(* IEC 61131-3 sources: SortJet_MasterSPS_Aufbau.fbsproj/09_Station/Shuttle/[101,102] Shuttle, 9 files *)

(* ---- Dickenverstellung_FB_V01_00_00.fb.st ---- *)
(* METADATA
{
	"v3Meta": {
		"objectGuid": "d815e3f2-dcd5-4a25-9c13-c3ee247e2cce"
	}
}
*)
FUNCTION_BLOCK Dickenverstellung_FB_V01_00_00
VAR_INPUT

  // BOOLEAN
  bpAktivieren                                   : BOOL; // Hinweis: Baustein aktivieren
  bpReset                                        : BOOL;
  bpStartePositionierung                         : BOOL;
  bpReferenz                                     : BOOL;
  bpFreigabe                                     : BOOL;
  bpOptionMotorischAktivieren                    : BOOL;
  bpOptionPneumatikAktivieren                    : BOOL;
  bpOption3WegeLogikDrehen                       : BOOL;
  bpOptionRollenleisteSchuetzSchaltungAktivieren : BOOL;
  bpOptionGegenhalterSchuetzSchaltungAktivieren  : BOOL;

  // ENUM
  epSollStellung : PneumatikZylinderStatus_EN;

  // STRUCT
  stStationsNummern  : Station_ST;

  // POINTER
  ppAntriebsInformationen : REFERENCE TO AntriebsInformationen;
  ppParameterBaustein     : REFERENCE TO Parameter_Dickenverstellung;  // Zeiger auf Parameterfeld

END_VAR
VAR_OUTPUT

  // BOOLEAN
  bpFehler                  : BOOL;
  bpDone                    : BOOL;
  bpResourceAktiv           : BOOL;
  bpInReferenz              : BOOL; // Status: Baustein/Antrieb ist referenziert

  // WORD
  wpFehlerNr : Fehlerkonstanten_EN;

  // ENUM
  eStatusStellung : PneumatikZylinderStatus_EN;

END_VAR
VAR

  // BOOLEAN
  blErsterZyklus   : BOOL := TRUE;

  // REAL
  rlZielPosition   : REAL;

  // TIMER
  tonlEndschalterFreifahren              : TON; // EINSCHALTVERZOEGERUNG:
  tonlWarteSchrittEndschalterFreifahren  : TON; // EINSCHALTVERZOEGERUNG:
  tonlMaxWarteAufResetErfolgreich        : TON; // EINSCHALTVERZOEGERUNG:
  tofHardwareEndschalterFrei             : TOF; // AUSSCHALTVERZOEGERUNG:
  toflAutoAbschaltung                    : TOF; // AUSSCHALTVERZOEGERUNG:

  // STEPS
  steplPositionieren    : Steps_TE;
  steplReferenz         : Steps_TE;
  steplReset            : Steps_TE;

  // Antrieb
  Antrieb : REFERENCE TO Rexroth_ctrlX_Drive_Eckelmann_MC_V01_02_02;

END_VAR
VAR_INPUT

  // HARDWARE EINGAENGE
  in_bEndschalterMax : BOOL; // Oeffner (TRUE = frei), gemappt; zum Umrichter ueber Signal-Steuerwort Bit 9, wirkt nur bei Endschalterquelle SPS

END_VAR
//-------------------------------------------------------------------------------------------------
// INITIALISIERUNG
//-------------------------------------------------------------------------------------------------
IF ( blErsterZyklus ) THEN

  IF ( __ISVALIDREF(ppAntriebsInformationen) ) THEN

    blErsterZyklus := FALSE;

    Antrieb REF= pgAntriebe[ppAntriebsInformationen.wAchsID];

    (* Hinweis:
       - Initialisierung Antriebsinformationen
    *)
    Antrieb.ppAntriebsInformationen REF= ppAntriebsInformationen;

    (* Hinweis:
       - Für die Zielpunktkontrolle muss im ersten Zyklus die Zielposition initialisiert werden
    *)
    Antrieb.rpZielPosition := Antrieb.rpIstPosition;

    (* Hinweis:
       - Antriebswerte vorinitialisieren
    *)
    Antrieb.rpGeschwindigkeit := ppAntriebsInformationen.rpMaxGeschwindigkeit;
    Antrieb.rpBeschleunigung  := ppAntriebsInformationen.rpMaxBeschleunigung;
    Antrieb.rpVerzoegerung    := ppAntriebsInformationen.rpMaxVerzoegerung;
    Antrieb.rpRuckzeit        := ppAntriebsInformationen.rpMaxRuckzeit;

  ELSE
    RETURN;
  END_IF

END_IF

// Endschalter zyklisch an den Antrieb geben, auch bei deaktivierter Bewegung
Antrieb.bpEndschalterMaxExtern := in_bEndschalterMax;

//-------------------------------------------------------------------------------------------------
// BAUSTEIN: AUSFUEHRUNG
//-------------------------------------------------------------------------------------------------
(* Hinweis:
   - Aktionen
*)
IF ( bpReset AND bpAktivieren ) THEN

  Reset();

ELSE

  IF ( bpAktivieren ) THEN
    Positionieren();
    Referenz();
    Ausgaenge();

    (* Hinweis:
       - Abschaltung
    *)
    toflAutoAbschaltung( IN :=     bpStartePositionierung
                         OR bpReferenz,
                         PT:= tgZeitAutoabschaltungEnergiesparModus );

    Antrieb.bpFreigabe := toflAutoAbschaltung.Q
                          AND bpAktivieren
                          AND bpFreigabe;

    Antrieb.rpRuckzeit := ppAntriebsInformationen.rpMaxRuckzeit;

    Antrieb.stStationsNummern := stStationsNummern;

  ELSE
    bpDone   := TRUE;
    bpFehler := FALSE;
    bpInReferenz := TRUE;

    eStatusStellung := epSollStellung;

    wpFehlerNr := cMELDUNG_NULL;

  END_IF // => bpAktiv

END_IF// => bpReset
END_FUNCTION_BLOCK

(* ---- Dickenverstellung_Schuetz_FB_V01_00_00.fb.st ---- *)
(* METADATA
{
	"v3Meta": {
		"objectGuid": "2c7452d1-eabd-4c4a-95fd-5aca04df1ee1"
	}
}
*)
FUNCTION_BLOCK Dickenverstellung_Schuetz_FB_V01_00_00
VAR_INPUT

  // BOOL
  bpAktivieren               : BOOL;
  bpVerstellungOeffnen       : BOOL;
  bpVerstellungSchliessen    : BOOL;
  bpReset                    : BOOL;

END_VAR
VAR_OUTPUT

  // BOOL
  bpFehler        : BOOL;
  bpDone          : BOOL;
  bpResourceAktiv : BOOL;

  // WORD
  wpFehlerNr      : Fehlerkonstanten_EN;

END_VAR

VAR

  // BOOL
  blErsterZyklus        : BOOL := TRUE;

  // TIMER
  tonlMaxWarteZeit                        : TON;
  tonlAntriebOK                           : TON;
  tonlMaximaleWartezeitAufReset           : TON;
  tonlFehlermeldungUnterdrueckenAntriebOK : TON;

  // STEPS
  steplVerstellungOeffnen      : Steps_TE;
  steplVerstellungSchliessen   : Steps_TE;
  steplReset                   : Steps_TE;

END_VAR

VAR
  // HARDWARE EINGÄNGE
  in_bVerstellungGeoeffnet         AT %I* : BOOL;
  in_bVerstellungGeschlossen       AT %I* : BOOL;
  in_bMotorstarter_OK              AT %I* : BOOL; // Sicherung des Kippantriebs ÖFFNER KONTAKT !!
  in_bBremseOK                     AT %I* : BOOL; // Sicherung des Kippantriebs ÖFFNER KONTAKT !!
  in_bSicherungMotorOK             AT %I* : BOOL;

  // HARDWARE AUSGÄNGE
  out_bVerstellungSchliessen       AT %Q* : BOOL;
  out_bVerstellungOeffnen          AT %Q* : BOOL;
  out_bBremseOeffnen               AT %Q* : BOOL;
  out_bMotorstarterReset           AT %Q* : BOOL;

END_VAR

//-------------------------------------------------------------------------------------------------
// BAUSTEIN: INITIALISIERUNG
//-------------------------------------------------------------------------------------------------
IF ( blErsterZyklus ) THEN
  blErsterZyklus := FALSE;

  (* Hinweis:
     - Timer initialisieren
  *)
  tonlAntriebOK(IN:=TRUE);
  tonlMaxWarteZeit(IN:=FALSE);
  tonlFehlermeldungUnterdrueckenAntriebOK( IN := FALSE );

END_IF

//-------------------------------------------------------------------------------------------------
// BAUSTEIN: AKTIONEN
//-------------------------------------------------------------------------------------------------
(* Hinweis:
   - Aktionen
*)
IF ( bpReset ) THEN

  bpReset                 := FALSE;
  bpVerstellungOeffnen    := FALSE;
  bpVerstellungSchliessen := FALSE;

  bpFehler        := FALSE;
  bpDone          := FALSE;
  bpResourceAktiv := FALSE;

  wpFehlerNr := cMELDUNG_NULL;

  out_bVerstellungSchliessen  := FALSE;
  out_bVerstellungOeffnen := FALSE;

ELSE

  IF ( bpAktivieren ) THEN

    VerstellungSchliessen();
    VerstellungOeffnen();

    out_bBremseOeffnen := out_bVerstellungOeffnen OR out_bVerstellungSchliessen;

    Meldungen();
    Timer();

  ELSE

    bpDone   := TRUE;
    bpFehler := FALSE;

  END_IF // => bpAktiv

END_IF// => bpReset
END_FUNCTION_BLOCK

(* ---- Greiferzange_FB_V01_00_00.fb.st ---- *)
(* METADATA
{
	"v3Meta": {
		"objectGuid": "50b45b59-5893-4c9c-b524-1732205d1fb3"
	}
}
*)
FUNCTION_BLOCK Greiferzange_FB_V01_00_00
VAR_INPUT

  // BOOLEAN
  bpReset                     : BOOL;
  bpAktivieren                : BOOL;
  bpFreigabe                  : BOOL; // FREIGABE Pneumatik: ohne Freigabe Ventile aus, Bewegung pausiert (Startbefehl bleibt erhalten)
  bpStartZylinderBewegung     : BOOL; // BETRIEBTYP: Greiferzange in die Soll-Stellung bewegen
  bpZylinderAbfragenVorhanden : BOOL := FALSE; // Hinweis: Endlagenabfragen der Zylinder vorhanden

  // TIME
  tpBewegungszeit             : TIME := T#700MS; // Bewegungszeit je Stellung ohne Abfragen bzw. beim Schliessen auf Glas

  // ENUM
  epSollZylinderStellung      : PneumatikZylinderStatus_EN; // eZylinderGeschlossen, eZylinderStellung16mm, eZylinderStellung23mm, eZylinderStellung29mm

END_VAR
VAR_OUTPUT

  // BOOLEAN
  bpFehler                    : BOOL;
  bpDone                      : BOOL;

  // WORD
  wpFehlerNr                  : Fehlerkonstanten_EN;

  // ENUM
  epStatusZylinderStellung    : PneumatikZylinderStatus_EN;

END_VAR
VAR

  // STEPS
  steplZylinderStellung       : Steps_TE;

  // TIMER
  tonlUeberwachungStellung      : TON; // EINSCHALTVERZOEGERUNG: Ueberwachung der Soll-Stellung mit Abfragen
  tonlWartezeitZylinderStellung : TON; // EINSCHALTVERZOEGERUNG: Bewegungszeit ohne Abfragen

END_VAR
VAR

  // HARDWARE EINGAENGE
  in_bStatusZylinder_Alle_Eingefahren AT %I* : BOOL; // STATUS: Zylinderabfrage [Eingefahren] Zange geschlossen
  in_bStatusZylinder_1_Ausgefahren    AT %I* : BOOL; // STATUS: Zylinderabfrage [Ausgefahren] Oeffnung 16 mm
  in_bStatusZylinder_2_Ausgefahren    AT %I* : BOOL; // STATUS: Zylinderabfrage [Ausgefahren] Oeffnung 23 mm
  in_bStatusZylinder_3_Ausgefahren    AT %I* : BOOL; // STATUS: Zylinderabfrage [Ausgefahren] Oeffnung 29 mm

  // HARDWARE AUSGAENGE
  out_bZylinder_1_Einfahren           AT %Q* : BOOL; // Impuls Zylinder 1 einfahren
  out_bZylinder_2_Einfahren           AT %Q* : BOOL; // Impuls Zylinder 2 einfahren
  out_bZylinder_3_Einfahren           AT %Q* : BOOL; // Impuls Zylinder 3 einfahren
  out_bZylinder_1_Ausfahren           AT %Q* : BOOL; // Impuls Zylinder 1 ausfahren [16 mm]
  out_bZylinder_2_Ausfahren           AT %Q* : BOOL; // Impuls Zylinder 2 ausfahren [23 mm]
  out_bZylinder_3_Ausfahren           AT %Q* : BOOL; // Impuls Zylinder 3 ausfahren [29 mm]

END_VAR
VAR CONSTANT

  // TIME
  cZEIT_UEBERWACHUNG_STELLUNG : TIME := T#5S;

END_VAR
(* Anmerkung:
   - Greiferzange mit drei Zylindern: geschlossen, Oeffnung 16 mm, 23 mm oder 29 mm
   - Vor dem Oeffnen werden alle Zylinder eingefahren, danach faehrt der Zylinder der Soll-Oeffnung aus
*)
//-------------------------------------------------------------------------------------------------
// BAUSTEIN: RESET / DEAKTIVIERT
//-------------------------------------------------------------------------------------------------
(* Hinweis:
   - Reset oder deaktiviert: Ausgaenge aus, Kette und Timer zuruecksetzen, Done und Fehler loeschen
   - Der Baustein setzt bpReset selbst zurueck, der Aufrufer wartet nicht auf Done
   - Ein deaktivierter Baustein meldet kein Done; der Aufrufer verknuepft das Warten auf Done
     mit der Aktivierung aus der MK (z.B. Greiferzange.bpDone OR NOT stStationsAufbau.bGreifer[wWand])
*)
IF ( bpReset OR NOT bpAktivieren ) THEN

  out_bZylinder_1_Einfahren := FALSE;
  out_bZylinder_2_Einfahren := FALSE;
  out_bZylinder_3_Einfahren := FALSE;
  out_bZylinder_1_Ausfahren := FALSE;
  out_bZylinder_2_Ausfahren := FALSE;
  out_bZylinder_3_Ausfahren := FALSE;

  bpStartZylinderBewegung := FALSE;

  steplZylinderStellung := STEP_0_E;

  tonlUeberwachungStellung( IN := FALSE );
  tonlWartezeitZylinderStellung( IN := FALSE );

  bpDone     := FALSE;
  bpFehler   := FALSE;
  wpFehlerNr := cMELDUNG_NULL;

  bpReset := FALSE;

  RETURN;

END_IF

//-------------------------------------------------------------------------------------------------
// BAUSTEIN: AKTIONEN
//-------------------------------------------------------------------------------------------------
(* Hinweis Freigabe Pneumatik:
   - Ohne Freigabe: Ventile aus, Kette und Ueberwachungszeiten zuruecksetzen (kein Timeout-Fehler)
   - Der Startbefehl bleibt erhalten: kommt die Freigabe zurueck, wird die Bewegung neu gestartet
*)
IF NOT bpFreigabe THEN
  out_bZylinder_1_Einfahren := FALSE;
  out_bZylinder_2_Einfahren := FALSE;
  out_bZylinder_3_Einfahren := FALSE;
  out_bZylinder_1_Ausfahren := FALSE;
  out_bZylinder_2_Ausfahren := FALSE;
  out_bZylinder_3_Ausfahren := FALSE;
  steplZylinderStellung := STEP_0_E;
  tonlUeberwachungStellung( IN := FALSE );
  tonlWartezeitZylinderStellung( IN := FALSE );
  bpDone := FALSE;
ELSE
  ZylinderBewegung();
END_IF

//-------------------------------------------------------------------------------------------------
// STATUS DER ZYLINDER
//-------------------------------------------------------------------------------------------------
(* Hinweis:
   - Status aus der Sensorik, wenn Abfragen vorhanden sind
   - Ohne Abfragen bleibt der Status, den die Schrittkette nach der Bewegungszeit setzt
*)
IF ( bpZylinderAbfragenVorhanden ) THEN

  IF ( in_bStatusZylinder_3_Ausgefahren ) THEN
    epStatusZylinderStellung := eZylinderStellung29mm;

  ELSIF ( in_bStatusZylinder_2_Ausgefahren ) THEN
    epStatusZylinderStellung := eZylinderStellung23mm;

  ELSIF ( in_bStatusZylinder_1_Ausgefahren ) THEN
    epStatusZylinderStellung := eZylinderStellung16mm;

  ELSIF ( in_bStatusZylinder_Alle_Eingefahren ) THEN
    epStatusZylinderStellung := eZylinderGeschlossen;

  ELSE
    epStatusZylinderStellung := eZylinderUndefiniert;

  END_IF

END_IF
END_FUNCTION_BLOCK

(* ---- Shuttle_FB_V01_00_00.fb.st ---- *)
(* METADATA
{
	"v3Meta": {
		"objectGuid": "a8175c8a-0e5e-42c5-a90c-c5e1a843dc34"
	}
}
*)
FUNCTION_BLOCK Shuttle_FB_V01_00_00
VAR_IN_OUT

  // STRUKT
  BasisStationsParameter : StationBasisParameter_ST;

END_VAR
VAR_INPUT

  // BOOLEAN
  bpShuttleAnhalten                      : BOOL; // HINWEIS: Nehmen der Verfahrfreigabe wenn bei der Folge- bzw. Nachfolgestation der Einlauf- / Auslauf- Sensor belegt wurde
  bpStarteFaecherwagensuche              : BOOL; // Der Fächerwagen kann mittels Sensor gesucht werden um die Fachpositionen zu bestimmen

  // WORD
  rpMinPosSwEsEingrenzung                : REAL;
  rpMaxPosSwEsEingrenzung                : REAL;

END_VAR
VAR_OUTPUT

  // BOOLEAN
  bpFaecherwagenGefunden                 : BOOL;

  // REAL
  rpAktuelleFaecherwagenPosition         : REAL;

  // DWORD
  dwpHandfunktionenReturn                : DWORD; // Aktive Handfunktionen, gleiche Bitbelegung wie dwlHandfunktionen

END_VAR
VAR

  // BOOL
  blErsterZyklus                         : BOOL := TRUE;// Initialisierungsphase
  blGeblaeseAktiv                        : BOOL;
  blBetriebsartHand                      : BOOL;
  blBetriebsartReset                     : BOOL;
  blBetriebartCheck                      : BOOL;
  blBetriebsartAutomatik                 : BOOL;
  blBetriebsartReferenz                  : BOOL;
  ablZielPositionErreicht                : ARRAY[cWAND_1..cANZAHL_WAENDE] OF BOOL; // Je Wand: Zielposition aus dem Auftrag der Wand stimmt mit der aktuellen Position ueberein [Toleranz rgMKZielPositionToleranz]
  blVorAbAuftragAktiv                    : ARRAY [cWAND_1..cANZAHL_WAENDE] OF BOOL; // STATUS: Merker ob die Komponenten Ansteuerung aktiv ist [Angesteuert mit dem Starten der Querfahrt](Autark gesteuert)
  blUpdateTimer                          : BOOL;
  blNachSystemcheckMerker                : BOOL; // Merkt sich, wenn der Systemcheck erfolgreich durchgeführt wurde, damit die Gebläse nicht nach dem Systemcheck ausgehen
  ablVortransportAktiv                   : ARRAY [cWAND_1..cANZAHL_WAENDE] OF BOOL; // STATUS: Merker ob der Vortransport (Autark gesteuert) aktiv ist -> Wichtig für den Austransport zum sicherstellen das erst dann Transportiert werden kann
  blDatenlichtschrankeUnterbrochenMelden : BOOL;
  blFehlerAusAutomatikBetrieb            : BOOL;
  blShuttleErreichbar                    : BOOL;
  blMerkerAuftragAktiv                   : BOOL;
  blMerkerEinOderAustransportAktiv       : BOOL;

  // WORD
  wlBetriebsart              : WORD;
  wlWatchIONachrichtenNummer : WORD;
  wlIndex                    : WORD;

  // DWORD
  dwlHandfunktionen                : DWORD;  // Handfunktionen: 0..31 Bit
  dwlHandfunktionenZuletztGesendet : DWORD;  // Rueckmeldung der Handfunktionen zum MMI

  // REAL
  rlLetztePosition  : REAL;

  // TIMER
  tonlMaxWarteAufResetErfolgreich       : TON;
  tonlUpdateTimer                       : TON; // Verfahrlogik
  tonWaitTimerAnsteuerungResourcen      : ARRAY[cWAND_1..cANZAHL_WAENDE] OF TON;
  tonWaitTimerAnsteuerungResourcenDone  : ARRAY[cWAND_1..cANZAHL_WAENDE] OF TON;

  toflGeblaeseHandfahren                : ARRAY[cWAND_1..cANZAHL_WAENDE] OF TOF;
  atoflSensorEinlauf                    : ARRAY[cWAND_1..cANZAHL_WAENDE] OF TOF;
  atoflSensorAuslauf                    : ARRAY[cWAND_1..cANZAHL_WAENDE] OF TOF;
  atoflSensorAUslaufStopp               : ARRAY[cWAND_1..cANZAHL_WAENDE] OF TOF;
  atoflSensorEinlaufStopp               : ARRAY[cWAND_1..cANZAHL_WAENDE] OF TOF;

  // TRIGGER
  rtlAutomatikActiv                     : R_TRIG;
  rtlGlastransportVerfahrfreigabe       : ARRAY [cWAND_1..cANZAHL_WAENDE] OF R_TRIG;
  rtlDatenlichtschrankeUnterbrochen     : R_TRIG;
  rtlFehlerMeldungGenerierenHandbetrieb : R_TRIG;
  rtlFehlerAusgeloestImAutomatikbetrieb : R_TRIG;
  artlVerfahrabbruchSensorik            : ARRAY [cWAND_1..cANZAHL_WAENDE] OF R_TRIG;
  artlWandverstellungPositionieren      : ARRAY [cWAND_1..cANZAHL_WAENDE] OF R_TRIG;
  rtlRackPositionGefunden               : R_TRIG;
  ftlBausteinDeaktivierung              : F_TRIG;

  // STEPS
  steplCheck                       : STEPS_TE;
  steplResetAntrieb                : STEPS_TE;
  steplReferenz                    : Steps_TE;
  steplVorabpositionierung         : STEPS_TE;
  steplFaecherwagensuche           : STEPS_TE;

  // BAUSTEINE
  Querfahrt                       : Querfahrt_Shuttle_FB_V01_00_00;
  Zentralschmierung               : Zentralschmierung_DLS_4xxi_FB_V01_00_00;
  Glastransport                   : ARRAY[cWAND_1..cANZAHL_WAENDE] OF Shuttle_Glastransport_FB_V01_00_00;
  Geblaese                        : ARRAY[cWAND_1..cANZAHL_WAENDE] OF Geblaese_Schuetz_FB_V01_00_00;
  Wandverstellung                 : ARRAY[cWAND_1..cANZAHL_WAENDE] OF Dickenverstellung_FB_V01_00_00;
  Kippen                          : Shuttle_Kippen_V01_00_00;

  Eintransport                    : ARRAY[cWAND_1..cANZAHL_WAENDE] OF Shuttle_Eintransport_FB_V01_00_00;
  Austransport                    : ARRAY[cWAND_1..cANZAHL_WAENDE] OF Shuttle_Austransport_FB_V01_00_00;
  Durchtransport                  : ARRAY[cWAND_1..cANZAHL_WAENDE] OF Shuttle_Durchtransport_FB_V01_00_00;
  AnsteuerungRessourcen           : ARRAY[cWAND_1..cANZAHL_WAENDE] OF Shuttle_Ansteuerung_Ressourcen_FB_V01_00_00;
  Greifer                         : ARRAY[cWAND_1..cANZAHL_WAENDE] OF Shuttle_Greifer_FB_V01_00_00; // Ausbaustufe stStationsAufbau.bGreifer

END_VAR
VAR
  // Alle Sensoren
  blAlleEinlaufStoppSensoren : BOOL; // wirksame Einlauf-Stopp-Sensoren (ohne MK: Einlaufsensor)
  blAlleAuslaufStoppSensoren : BOOL;
  ablSensorEinlaufStopp      : ARRAY[cWAND_1..cANZAHL_WAENDE] OF BOOL; // wirksamer Einlauf-Stopp-Sensor (ohne MK: Einlaufsensor)
  ablSensorAuslaufStopp      : ARRAY[cWAND_1..cANZAHL_WAENDE] OF BOOL; // wirksamer Auslauf-Stopp-Sensor (ohne MK: Auslaufsensor)
  blAlleVerfahrfreigaben     : BOOL;
  blAlleGreiferSicher        : BOOL; // Alle Greifer in sicherer Position mit eingefahrenen Glasrueckhaltern (oder nicht vorhanden)
  blGreiferVor               : BOOL; // Handbetrieb Greifer: Taster MMI oder Visu (Aktion Handfunktionen)
  blGreiferZurueck           : BOOL;
  blGreiferReferenz          : BOOL;
  blGreiferAusfahren         : BOOL;
  blGreiferEinfahren         : BOOL;
  ablQuittScheibe            : ARRAY[cWAND_1..cANZAHL_WAENDE] OF BOOL; // Scheibenquittierung Glastransport bzw. Greifer
  blDone                     : BOOL;
  blFehlerAktiv              : BOOL;

  // HARDWARE EINGAENGE
  in_bSensorEinlauf                                   : ARRAY[cWAND_1..cANZAHL_WAENDE] OF BOOL; // Shuttle Sensoren von links nach rechts Sensor 1
  in_bSensorAuslauf                                   : ARRAY[cWAND_1..cANZAHL_WAENDE] OF BOOL; // Shuttle Sensoren von links nach rechts Sensor 4
  in_bSensorEinlaufVorab                              : ARRAY[cWAND_1..cANZAHL_WAENDE] OF BOOL; // Shuttle Sensoren von links nach rechts Sensor 2
  in_bSensorAuslaufVorab                              : ARRAY[cWAND_1..cANZAHL_WAENDE] OF BOOL; // Shuttle Sensoren von links nach rechts Sensor 3
  in_bSensorEinlaufStopp                              : ARRAY[cWAND_1..cANZAHL_WAENDE] OF BOOL; // Shuttle Sensoren von links nach rechts Sensor 0 (nur mit MK bSensorEinlaufStopp)
  in_bSensorAuslaufStopp                              : ARRAY[cWAND_1..cANZAHL_WAENDE] OF BOOL; // Shuttle Sensoren von links nach rechts Sensor 5 (nur mit MK bSensorAuslaufStopp)
  in_bDatenlichtschrankeShuttlebahnOK          AT %I* : BOOL; // Bauteil an der Shuttlebahn => Sender / Empfaenger
  in_bDatenlichtschrankeShuttleOK              AT %I* : BOOL; // Bauteil auf dem Shuttle => Sender / Empfaenger
  in_bNetzteil_24V_OK                          AT %I* : BOOL;
  in_bKlimageraet_OK                                  : BOOL;
  in_bSicherungen24V_OK                               : BOOL;
  in_bDruckluft_OK                             AT %I* : BOOL;
  in_bSicherungKompressor_OK                   AT %I* : BOOL;
  in_bLSQuerfahrtBremseOK                      AT %I* : BOOL;

  in_bSicherungen230V_OK                       AT %I* : BOOL;
  in_iAnalogwertChannel1                              : INT; // Hinweis: Eingaenge des Analogmoduls u.a fuer die automatische Fachaufnahme
  in_iAnalogwertChannel2                              : INT; // Hinweis: Eingaenge des Analogmoduls u.a fuer die automatische Fachaufnahme
  in_bWandverstellungsAntriebsSicherungOK      AT %I* : BOOL;
  in_bWandverstellungsBremsSicherungOK         AT %I* : BOOL;
  in_bFaecherwagenSuchSensor                          : BOOL; // Shuttle Sensor zum Suchen der Fächerwagen um die Fachpositionen zu bestimmen

  aHand : ARRAY[0..31] OF BOOL;
  i     : INT;

END_VAR
VAR CONSTANT

  // TIME
  ZEIT_SENSOR_ENTPRELLEN         : TIME := T#50ms;

END_VAR
(* Anmerkung:
   - Shuttle Koordinationsbaustein regelt das komplette Shuttle
*)
//-------------------------------------------------------------------------------------------------
// BAUSTEIN: INITIALISIERUNG
//-------------------------------------------------------------------------------------------------

IF ( blErsterZyklus ) THEN
  blErsterZyklus:=FALSE;

  (* Wichtig:
     - Initialisierung
  *)
  A_Baustein_Initialisierung();

END_IF

FOR wlIndex := cWAND_1 TO cANZAHL_WAENDE DO
  in_bSensorEinlauf[wlIndex] := Glastransport[wlIndex].Antrieb.udipEingaengeUmrichter.cXG31_1_I_1;
  in_bSensorAuslauf[wlIndex] := Glastransport[wlIndex].Antrieb.udipEingaengeUmrichter.cXG31_2_I_2;

  ablSensorEinlaufStopp[wlIndex] := SEL( BasisStationsParameter.stMKs.stStationsAufbau.bSensorEinlaufStopp, in_bSensorEinlauf[wlIndex], in_bSensorEinlaufStopp[wlIndex] );
  ablSensorAuslaufStopp[wlIndex] := SEL( BasisStationsParameter.stMKs.stStationsAufbau.bSensorAuslaufStopp, in_bSensorAuslauf[wlIndex], in_bSensorAuslaufStopp[wlIndex] );
END_FOR

blAlleEinlaufStoppSensoren := FALSE;
blAlleAuslaufStoppSensoren := FALSE;
blAlleVerfahrfreigaben     := TRUE;
blAlleGreiferSicher        := TRUE;

FOR wlIndex := cWAND_1 TO cANZAHL_WAENDE DO
  blAlleGreiferSicher        := blAlleGreiferSicher
                                AND (    ( Greifer[wlIndex].bpSicherePosition AND Greifer[wlIndex].bpGlasRueckhalterEingefahren )
                                      OR NOT BasisStationsParameter.stMKs.stStationsAufbau.bGreifer[wlIndex] );
  blAlleEinlaufStoppSensoren := blAlleEinlaufStoppSensoren OR ablSensorEinlaufStopp[wlIndex];
  blAlleAuslaufStoppSensoren := blAlleAuslaufStoppSensoren OR ablSensorAuslaufStopp[wlIndex];
  blAlleVerfahrfreigaben     := blAlleVerfahrfreigaben AND Glastransport[wlIndex].bpVerfahrFreigabe;
END_FOR

//-------------------------------------------------------------------------------------------------
// DEAKTIVIERUNG
//-------------------------------------------------------------------------------------------------

(* Hinweis:
   - Werte wieder passend abloeschen, wenn der Baustein wieder aktiviert wird
*)
ftlBausteinDeaktivierung( CLK := BasisStationsParameter.stMKs.bDeaktivieren );

IF ( ftlBausteinDeaktivierung.Q ) THEN

  SendShuttlePosition();

  FOR wlIndex := cWAND_1 TO cANZAHL_WAENDE DO
    BasisStationsParameter.bEintransportAbgeschlossen[wlIndex] := FALSE;
    BasisStationsParameter.bAustransportAbgeschlossen[wlIndex] := FALSE;
  END_FOR

  BasisStationsParameter.bIstReferenziert       := FALSE;
  BasisStationsParameter.bCheckAbgeschlossen    := FALSE;
  BasisStationsParameter.bReferenzAbgeschlossen := FALSE;

END_IF

(* Hinweis:
   - Deaktivierung des Bausteins
     => Der Baustein wird zum Ende der RETURN-Anweisung verlassen
*)
IF ( BasisStationsParameter.stMKs.bDeaktivieren ) THEN

  IF ( apgShuttleVerfahrparameter[BasisStationsParameter.stMKs.stStationsNummern.NummerSPS].eParkposition = PARKPOSITION_MAX ) THEN
    BasisStationsParameter.rAktuellePositionQuerfahrt := apgShuttleVerfahrparameter[BasisStationsParameter.stMKs.stStationsNummern.NummerSPS].rParkpositionMaximum;
  ELSE
    BasisStationsParameter.rAktuellePositionQuerfahrt := apgShuttleVerfahrparameter[BasisStationsParameter.stMKs.stStationsNummern.NummerSPS].rParkpositionMinimum;
  END_IF

  FOR wlIndex := cWAND_1 TO cANZAHL_WAENDE DO
    BasisStationsParameter.bEintransportAbgeschlossen[wlIndex] := TRUE;
    BasisStationsParameter.bAustransportAbgeschlossen[wlIndex] := TRUE;

    IF ( BasisStationsParameter.bCheck ) THEN

      IF BasisStationsParameter.stMKs.stStationsAufbau.bGlastransport[wlIndex] THEN
        rSps2MmiMessungScheibenlaenge   := 0;
        wSps2MmiMessungStationNummer    := BasisStationsParameter.stMKs.stStationsNummern.NummerIntern;
        wSps2MmiMessungSlotNummer       := wlIndex;
        iSps2MmiMessungScheibenanzahl   := 0;

        MsgToMmi( auftragsnr_w := SB0_SPS_SETSHEETSONSTATION );
      END_IF
    END_IF

  END_FOR

  BasisStationsParameter.bIstReferenziert       := TRUE;
  BasisStationsParameter.bCheckAbgeschlossen    := TRUE;
  BasisStationsParameter.bReferenzAbgeschlossen := TRUE;
  BasisStationsParameter.bReset                 := FALSE;

  BasisStationsParameter.bFehler       := FALSE;
  BasisStationsParameter.wFehlerNummer := cMELDUNG_NULL;

  HandfunktionenStatus();
  RETURN;

END_IF

//-------------------------------------------------------------------------------------------------
// AKTIONEN
//-------------------------------------------------------------------------------------------------
Betriebsart();

SystemCheck();

(* Hinweis:
   - Automatik-Aktionen
*)
FOR wlIndex := cWAND_1 TO cANZAHL_WAENDE DO
  Eintransport[wlIndex]( BasisStationsParameter := BasisStationsParameter,
                         wWand := wlIndex,
                         bpGeblaeseAktiv := Geblaese[wlIndex].bpDone,
                         bpAutomatikAktiv := BasisStationsParameter.bAutomatik,
                         bpVorAbAuftragAktiv := blVorAbAuftragAktiv[wlIndex],
                         bpZielPositionErreicht := ablZielPositionErreicht[wlIndex],
                         Glastransport := Glastransport[wlIndex],
                         Kippen := Kippen,
                         Wandverstellung := Wandverstellung[wlIndex],
                         Geblaese := Geblaese[wlIndex],
                         bpGreiferAktiv := BasisStationsParameter.stMKs.stStationsAufbau.bGreifer[wlIndex],
                         Greifer := Greifer[wlIndex]
                       );
  Austransport[wlIndex]( BasisStationsParameter := BasisStationsParameter,
                         wWand := wlIndex,
                         bpGeblaeseAktiv := Geblaese[wlIndex].bpDone,
                         bpAutomatikAktiv := BasisStationsParameter.bAutomatik,
                         bpVorAbAuftragAktiv := blVorAbAuftragAktiv[wlIndex],
                         bpZielPositionErreicht := ablZielPositionErreicht[wlIndex],
                         Glastransport := Glastransport[wlIndex],
                         Kippen := Kippen,
                         Wandverstellung := Wandverstellung[wlIndex],
                         Geblaese := Geblaese[wlIndex],
                         bpGreiferAktiv := BasisStationsParameter.stMKs.stStationsAufbau.bGreifer[wlIndex],
                         Greifer := Greifer[wlIndex]
                       );

  Durchtransport[wlIndex]( BasisStationsParameter := BasisStationsParameter,
                           wWand := wlIndex,
                           bpGeblaeseAktiv := Geblaese[wlIndex].bpDone,
                           bpAutomatikAktiv := BasisStationsParameter.bAutomatik,
                           bpVorAbAuftragAktiv := blVorAbAuftragAktiv[wlIndex],
                           bpZielPositionErreicht := ablZielPositionErreicht[wlIndex],
                           Glastransport := Glastransport[wlIndex],
                           Kippen := Kippen,
                           Wandverstellung := Wandverstellung[wlIndex],
                           Geblaese := Geblaese[wlIndex]
                         );
  AnsteuerungRessourcen[wlIndex]( BasisStationsParameter := BasisStationsParameter,
                                  wWand := wlIndex,
                                  bpGeblaeseAktiv := Geblaese[wlIndex].bpDone,
                                  bpAutomatikAktiv := BasisStationsParameter.bAutomatik,
                                  bpVorAbAuftragAktiv := blVorAbAuftragAktiv[wlIndex],
                                  bpZielPositionErreicht := ablZielPositionErreicht[wlIndex],
                                  Glastransport := Glastransport[wlIndex],
                                  Kippen := Kippen,
                                  Wandverstellung := Wandverstellung[wlIndex],
                                  Geblaese := Geblaese[wlIndex],
                                  bpGreiferAktiv := BasisStationsParameter.stMKs.stStationsAufbau.bGreifer[wlIndex],
                                  Greifer := Greifer[wlIndex]
                                );
END_FOR

Vorabpositionierung();

SensorenFreifahren();
FaecherwagenSuche();

(* Hinweis:
   - Basis-Aktionen
*)
Reset();
Referenz();
Meldungen();
Handfunktionen();

A_Geblaese();
A_Aufrufe();
A_Schnittstelle();
A_Ausgaenge();
END_FUNCTION_BLOCK

(* ---- Shuttle_Glastransport_FB_V01_00_00.fb.st ---- *)
(* METADATA
{
	"v3Meta": {
		"objectGuid": "bced77b5-e61c-4af0-a672-a0da8c7118bb"
	}
}
*)
FUNCTION_BLOCK Shuttle_Glastransport_FB_V01_00_00
VAR_INPUT

  bpDurchtransport                 : BOOL; // BETRIEBSMODUS[AUTOMATIK]: Eintransport-Schrittkette starten
  bpEintransport                   : BOOL; // BETRIEBSMODUS[AUTOMATIK]: Eintransport-Schrittkette starten
  bpRueckwaertsEintransportieren   : BOOL; // BETRIEBSMODUS[AUTOMATIK]: Eintransport Richtung -Rueckwaerts ueber den Auslaufsensor
  bpAustransport                   : BOOL; // BETRIEBSMODUS[AUTOMATIK]: Autransport-Schrittkette starten
  bpRueckwaertsAustransportieren   : BOOL; // BETRIEBSMODUS[AUTOMATIK]: Austransport Richtung -Rueckwaerts ueber den Einlaufsensor
  bpRueckwaertsSystemcheck         : BOOL;
  bpVortransport                   : BOOL; // BETRIEBSMODUS[AUTOMATIK]: Vortransport-Schrittkette starten
  bpVortransportRueck              : BOOL; // BETRIEBSMODUS[AUTOMATIK]: Vortransport-Schrittkette starten
  bpStarteSensorFreiFahren         : BOOL := FALSE; // BETRIEBSMODUS[AUTOMATIK]:
  bpHandfahrenPlus                 : BOOL; // BETRIEBSMODUS HANDBETRIEB: Im Handbetrieb den Riemen in positive Glasflussrichtung bewegen
  bpHandfahrenMinus                : BOOL; // BETRIEBSMODUS HANDBETRIEB: Im Handbetrieb den Riemen in negative Glasflussrichtung bewegen
  bpFahreReferenz                  : BOOL; // BETRIEBSMODUS: Antrieb referenzieren
  bpStarteVorabPositionierung      : BOOL; // BETRIEBSMODUS Positionieren der Scheibe fuer den Austransport
  bpStarteVorabPositionierungRueckwaertig : BOOL; // BETRIEBSMODUS Positionieren der Scheibe fuer den Austransport rueckwaerts (ueber den Einlaufsensor)
  bpCheck                          : BOOL;
  bpReset                          : BOOL;
  bpCheckMitVorgaenger             : BOOL; // Status: SystemCheck mit der Vorgaenger- Station
  bpCheckMitNachfolger             : BOOL; // Status: SystemCheck mit der Nachfolger- Station
  bpAutomatikAktiv                 : BOOL;
  bpFreigabe                       : BOOL; // Status: Der Riemen ist Freigegeben und kann Prozesse abarbeiten
  bpMessrichtungNegativ            : BOOL := FALSE; // HINWEIS: TRUE = Messrichtung negativ, FALSE = Messrichtung positiv
  bpAktivieren                     : BOOL := TRUE; // WICHTIG: Aktivieren des Bausteins
  bpScheibentrennung               : BOOL := FALSE;
  bpTransferstationTransfershuttle : BOOL := FALSE;
  bpSensorEinlauf                  : BOOL; // Sensoren von links nach rechts Sensor 1
  bpSensorEinlaufVorab             : BOOL; // Sensoren von links nach rechts Sensor 2
  bpSensorAuslaufVorab             : BOOL; // Sensoren von links nach rechts Sensor 3
  bpSensorAuslauf                  : BOOL; // Sensoren von links nach rechts Sensor 4
  bpSensorEinlaufStopp             : BOOL; // Sensoren von links nach rechts Sensor 0 (Verfahrfreigabe, Notbremse und Scheibe hat Shuttle verlassen im Rueckwaertstransport)
  bpSensorAuslaufStopp             : BOOL; // Sensoren von links nach rechts Sensor 5
  bpScheibeNachSystemcheckAufAuslaufsensor : BOOL;
  bpTeilnehmerErreichbar           : BOOL;
  bpMessungSystemCheckAktiv        : BOOL;
  bpSlaveAntriebVorhanden          : BOOL;

  // OPTIONEN
  bpOptionMasterSlaveTransport     : BOOL;

  // GREIFER
  bpStarteSlaveKopplungGreifer      : BOOL; // BETRIEBSMODUS GREIFER: Glastransport als Slave auf die Greiferachse koppeln
  bpStarteKorrekturfahrt            : BOOL; // BETRIEBSMODUS GREIFER: Sensor der Greiferseite frei fahren (uebergrosse Scheibe / nach dem Austransport)
  bpKorrekturfahrtRueckwaerts       : BOOL; // BETRIEBSMODUS GREIFER: TRUE = Auslaufsensor frei fahren, FALSE = Einlaufsensor frei fahren
  bpStarteGlasPositionierungGreifer : BOOL; // BETRIEBSMODUS GREIFER: Scheibe fuer den Austransport mit dem Greifer positionieren
  bpGlasPositionierungEinlaufseite  : BOOL; // BETRIEBSMODUS GREIFER: TRUE = ueber den Einlaufsensor positionieren, FALSE = ueber den Auslaufsensor
  wpAchsIDGreifer                   : WORD; // Achs-ID der Greiferachse (Master der Kopplung)
  rpWegGlasUebergabeposition        : REAL; // Weg der Scheibe ueber den Sensor der Greiferseite

  // WORD
  wpWandNr                    : WORD;

  // ENUM
  eStationsTyp                 : StationsTyp_EN; // Typ der Station [ Shuttle \ Station \ Faecherwagen \ etc. ]
  wpGlastyp                   : GlasTyp_EN; // AUFTRAGSDATEN : Unterscheidung fuer den Eintransports -> Grosse Scheiben

  // STRUCT
  InGlasTransportNachfolger   : Interface_GlasTransport; // STRUKTUR: Informationen ueber den Aus- Ein- Transport WAND 2
  InGlasTransportVorgaenger   : Interface_GlasTransport; // STRUKTUR: Informationen ueber den Aus- Ein- Transport WAND 2
  pAuftrag                    : Auftragsdaten_ST;        // AUFTRAG: Aktuelle daten zum Auftrag [Laenge, Hoehe, Modelle]
  stStationsNummern           : Station_ST;
  stMasterSlaveConfig         : MasterSlaveConfig_ST;

  // POINTER
  ppParameterBaustein           : REFERENCE TO Parameter_ShuttleGlastransport;
  ppAntriebsInformationen       : REFERENCE TO AntriebsInformationen;
  ppAntriebsInformationenSlave  : REFERENCE TO AntriebsInformationen;

END_VAR
VAR_OUTPUT

  // BOOLEAN
  bpDone                                      : BOOL;
  bpFehler                                    : BOOL;
  bprtScheibe                                 : BOOL;
  bpStationBelegt                             : BOOL;
  bpVerfahrFreigabe                           : BOOL;
  bpVortransportAktiv                         : BOOL; // STATUS: Merker ob der Vortransport (Autark gesteuert) aktiv ist -> Wichtig für den Austransport zum sicherstellen das erst dann Transportiert werden kann
  bpPositionierungAbgeschlossen               : BOOL; // HINWEIS:
  bpOutBereitZumAustransport                  : BOOL;
  bpOutBereitZumEintransport                  : BOOL;
  bpSlaveAktiv                                : BOOL; // STATUS: dem Baustein melden das der Slavebetrieb aktiv ist
  bpFreigabeQuerfahrt                         : BOOL; // HINWEIS: Freigabe setzen das die Querfahrt verfahren kann
  bpAuftragAktiv                              : BOOL;
  bpGreiferSlaveAktiv                         : BOOL; // STATUS: Glastransport ist auf die Greiferachse gekoppelt
  bpKorrekturfahrtAbgeschlossen               : BOOL; // STATUS: Korrekturfahrt fuer den Greifer abgeschlossen
  bpGlasPositionierungGreiferAbgeschlossen    : BOOL; // STATUS: Scheibe fuer den Greifer positioniert

  // WORD
  wpFehlerNr             : Fehlerkonstanten_EN;

  // DWORD
  dwpWartezeit              : DWORD :=0 ;// STATISTIK: Beschreibt die Zeit zwischen Anlegeauftrag und betaetigen des Tasters zum Eintransport

  // REAL
  rpOutGeschwindigkeit        : REAL;
  rlGlasgewicht               : REAL;

END_VAR
VAR

  // BOOLEAN
  blErsterZyklus                              : BOOL := TRUE;
  blSensorFreifahren                          : BOOL;
  blScheibenMerker                            : BOOL; // Merken da eien Scheibe den Auslaufsensor / Einlaufsensor beim Eintransport weiter
  blReduzierteGeschwindigkeit                 : BOOL;
  blAntriebsKopplungAktiv                     : BOOL;
  blStarteSlaveKopplung                       : BOOL;

  // INT
  ilScheibenZaehler  : INT;

  // REAL
  rlScheibenMessungErgebnis         : REAL; // SystemCheck
  rlAntriebIstPositionBeiStart      : REAL;
  rlMaxStreckeErsteScheibe          : REAL; // Max. Weg bis zur ersten Scheibe: Laenge der abgebenden Station, ohne bekannte Laenge die eigene Stationslaenge
  rlStreckeBisZurVerzoegerung       : REAL;
  rlPositionScheibenAnfangErkannt   : REAL;
  rlGeschwindigkeitEintransport     : REAL;
  rlGefahreneStreckeEintransport    : REAL; // Weg-Merker fuer die Strecke die beim Eintransport zurueck gelegt werden muss laut Auftrag

  // STEPS
  steplDurchtransport           : Steps_TE;
  steplEintransport             : Steps_TE;
  steplEintransportRueckwaertig : Steps_TE;
  steplAustransport             : Steps_TE;
  steplAustransportRueckwaertig : Steps_TE;
  steplSlave                    : Steps_TE;
  steplCheck                    : Steps_TE;
  steplReset                    : Steps_TE;
  steplReferenz                 : Steps_TE;
  steplVorabpositionieren       : STEPS_TE; // Hinweis: Positionierung ueber den Auslaufsensor
  steplVorabpositionierenRueckwaertig : STEPS_TE; // Hinweis: Positionierung ueber den Einlaufsensor
  steplSensorFreiFahren         : Steps_TE;
  steplVortransport             : Steps_TE;
  steplVortransportRueckwertig  : Steps_TE;
  steplSlaveGreifer             : Steps_TE;
  steplKorrekturfahrt           : Steps_TE;
  steplGlasPositionierungGreifer : Steps_TE;

  steplCheckMerker : Steps_TE;

  // TIMER
  toflAutoAbschaltung                : TOF; // AUSSCHALTVERZOEGERUNG:
  toflEinlaufsensor                  : TOF; // AUSSCHALTVERZOEGERUNG: Entprellen der Sensoren
  toflAuslaufsensor                  : TOF; // AUSSCHALTVERZOEGERUNG: Entprellen der Sensoren
  toflAuslaufsensorSTOP              : TOF; // AUSSCHALTVERZOEGERUNG: Entprellen der Sensoren
  toflEinlaufsensorSTOP              : TOF; // AUSSCHALTVERZOEGERUNG: Entprellen der Sensoren
  toflEinlaufsensorFrei              : TOF; // AUSSCHALTVERZOEGERUNG: Haelt die positive Flanke des Auslaufsensor eine gewissen Zeit aufrecht ( Freifahren des Sensors )
  toflAuslaufsensorFrei              : TOF; // AUSSCHALTVERZOEGERUNG: Haelt die positive Flanke des Auslaufsensor eine gewissen Zeit aufrecht ( Freifahren des Sensors )
  tonlMaxWarteAufResetErfolgreich    : TON; // EINSCHALTVERZOEGERUNG:
  tonlWarteSchritt                   : TON; // EINSCHALTVERZOEGERUNG:
  tonlAntriebNichtFreigegeben        : TON; // EINSCHALTVERZOEGERUNG:
  tonlUberwachungSlaveAktiv          : TON; // EINSCHALTVERZOEGERUNG:
  tonlSlaveKopplungDeaktiviert       : TON;
  tonlSlaveAntriebNichtFreigegeben   : TON; // Ueberwachung: Master/Slave nicht betriebsbereit
  tonlUeberwachungSlaveGreifer       : TON; // Ueberwachung: Kopplung auf die Greiferachse
  tonlUeberwachungGreiferBetrieb      : TON; // Ueberwachung: Antrieb bereit fuer Korrekturfahrt / Positionierung fuer den Greifer

  // TIME
  tlWarteZeiteAufnahme               : TIME; // STATISTIK: Zeit Ermittlung von evtl. Wartezeiten

  // STRING
  stlLogString    : STRING;

  // Antrieb
  Scheibenmessung  : Scheibenmessung_FB_V01_00_00;

  // Antrieb
  Antrieb       : REFERENCE TO Rexroth_ctrlX_Drive_Eckelmann_MC_V01_02_02;
  Antrieb_Slave : REFERENCE TO Rexroth_ctrlX_Drive_Eckelmann_MC_V01_02_02;

END_VAR
VAR CONSTANT

  // TIME
  cZEIT_UEBERWACHUNG_ANTRIEBSFREIGABE : TIME := T#5S;
  cUEBERWACHUNG_SLAVE_AKTIV           : TIME :=T#1S;

END_VAR

//-------------------------------------------------------------------------------------------------
// INITIALISIERUNG
//-------------------------------------------------------------------------------------------------
IF ( blErsterZyklus ) THEN

  IF ( __ISVALIDREF(ppAntriebsInformationen) ) THEN

    blErsterZyklus            := FALSE;

    Antrieb REF= pgAntriebe[ppAntriebsInformationen.wAchsID];
    IF ( __ISVALIDREF(ppAntriebsInformationenSlave) ) THEN
      Antrieb_Slave REF= pgAntriebe[ppAntriebsInformationenSlave.wAchsID];
    END_IF

    (* Hinweis:
       - Initialisierung Antriebsinformationen
    *)
    Antrieb.ppAntriebsInformationen REF= ppAntriebsInformationen;
    Antrieb.stStationsNummern := stStationsNummern;
    IF ( __ISVALIDREF(Antrieb_Slave) AND __ISVALIDREF(ppAntriebsInformationenSlave) ) THEN
      Antrieb_Slave.ppAntriebsInformationen REF= ppAntriebsInformationenSlave;
      Antrieb_Slave.stStationsNummern := stStationsNummern;
    END_IF

    (* Hinweis:
       - Antriebswerte vorinitialisieren
    *)
    Antrieb.rpGeschwindigkeit := ppAntriebsInformationen.rpMaxGeschwindigkeit;
    Antrieb.rpBeschleunigung  := ppAntriebsInformationen.rpMaxBeschleunigung;
    Antrieb.rpVerzoegerung    := ppAntriebsInformationen.rpMaxVerzoegerung;
    Antrieb.rpRuckzeit        := ppAntriebsInformationen.rpMaxRuckzeit;

    (* Hinweis:
       - Antriebswerte vorinitialisieren
    *)
    IF ( __ISVALIDREF(Antrieb_Slave) AND __ISVALIDREF(ppAntriebsInformationenSlave) ) THEN
      Antrieb_Slave.rpGeschwindigkeit := REAL#0;
      Antrieb_Slave.rpBeschleunigung  := ppAntriebsInformationenSlave.rpMaxBeschleunigung;
      Antrieb_Slave.rpVerzoegerung    := ppAntriebsInformationenSlave.rpMaxVerzoegerung;
      Antrieb_Slave.rpRuckzeit        := ppAntriebsInformationenSlave.rpMaxRuckzeit;
    END_IF

    // Pointer
    //   - Initialisierung zur vermeidung von null Pointerexceptions
    //     => Scheibenmessung
    Scheibenmessung.ppAntriebsInformationen REF= ppAntriebsInformationen;
    Scheibenmessung.ppAntrieb               REF= Antrieb;
    Scheibenmessung.pbpVorstopSensor        REF= bgFALSE;
    Scheibenmessung.pbpEinlaufSensor        REF= bgFALSE;

  ELSE
    RETURN;
  END_IF

END_IF

//-------------------------------------------------------------------------------------------------
// DEAKTIVIEREN
//-------------------------------------------------------------------------------------------------
IF ( NOT bpAktivieren ) THEN

  bpVerfahrFreigabe := TRUE;
  bpDone := TRUE;

  (* Hinweis:
     - Ausnahmesituationen
  *)
  bpFehler   := FALSE;
  wpFehlerNr := cMELDUNG_NULL;

  RETURN;

END_IF

//-------------------------------------------------------------------------------------------------
// TIMER, EINSTELLUNGEN, ETC.
//-------------------------------------------------------------------------------------------------
(* Hinweis:
   - Sensorenflackern
*)
toflEinlaufsensor(IN := bpSensorEinlauf, PT := t#50ms);
toflAuslaufsensor(IN := bpSensorAuslauf, PT := t#50ms);
toflAuslaufsensorSTOP(IN := bpSensorAuslaufStopp, PT := t#50ms);
toflEinlaufsensorSTOP(IN := bpSensorEinlaufStopp, PT := t#50ms);

// TIMER:
//   - Sensorenflackern
//     => Haelt die positive Flanke des Auslaufsensor eine gewissen Zeit aufrecht ( Freifahren des Sensors )
toflAuslaufsensorFrei(IN := bpSensorAuslauf, PT := t#100ms);
toflEinlaufsensorFrei(IN := bpSensorEinlauf, PT := t#100ms);

//-------------------------------------------------------------------------------------------------
// AKTIONEN
//-------------------------------------------------------------------------------------------------

(* Hinweis:
   - SystemCheck - Aktion
*)
SystemCheck();

(* Hinweis:
   - SystemCheck - Aktion
*)
Eintransport();
Eintransport_Rueckwertig();

Durchtransport();

Austransport();
Austransport_Rueckwertig();

GlasVorabPositionierung();
GlasVorabPositionierung_Rueckwaertig();

CASE eStationsTyp OF

  eInputShuttle:
    Vortransport_Inputshuttle();
    Vortransport_Rueckwertig();

  eOutputShuttle:
    Vortransport();
    Vortransport_Rueckwertig();

END_CASE

SensorenFreifahren();

(* Hinweis:
   - Zusammenspiel mit dem Shuttle-Greifer (nur mit stStationsAufbau.bGreifer angefordert)
*)
GlasPositionierungGreifer();
Korrekturfahrt();
SlaveBetriebGreifer();

IF ( bpSlaveAntriebVorhanden ) THEN
  Slave_Antrieb();
ELSE
  blAntriebsKopplungAktiv := TRUE;
END_IF
(* Hinweis:
   - Basis- Aktionen
*)
Reset();
Referenz();
Meldungen();
Handfunktionen();
Ausgaenge();

//-------------------------------------------------------------------------------------------------
// FREIGABEN UND BAUSTEINAUFRUFE
//-------------------------------------------------------------------------------------------------
(* Hinweis:
   - Freigaben des ANtriebs
*)
toflAutoAbschaltung( IN := (  bpAutomatikAktiv
                             AND ( bpEintransport
                                   OR bpRueckwaertsEintransportieren
                                   OR bpDurchtransport
                                   OR bpVortransport
                                   OR bpVortransportRueck
                                   OR bpAustransport
                                   OR bpRueckwaertsAustransportieren
                                   OR bpStarteSensorFreiFahren
                                   OR bpStarteVorabPositionierung
                                   OR bpStarteVorabPositionierungRueckwaertig
                                   OR bpStarteSlaveKopplungGreifer
                                   OR bpStarteKorrekturfahrt
                                   OR bpStarteGlasPositionierungGreifer ) )
                     OR bpCheck
                     OR bpHandfahrenMinus
                     OR bpHandfahrenPlus
                     OR bpFahreReferenz
                     OR bpStarteSlaveKopplungGreifer
                     OR blStarteSlaveKopplung,
                     PT:= tgZeitAutoabschaltungEnergiesparModus );

// Aufruf Antrieb
Antrieb.bpFreigabe        := toflAutoAbschaltung.Q AND bpFreigabe;
Antrieb.stStationsNummern := stStationsNummern;
Antrieb.rpRuckzeit        := ppAntriebsInformationen.rpMaxRuckzeit;

Antrieb_Slave.bpFreigabe        := toflAutoAbschaltung.Q AND bpFreigabe;
Antrieb_Slave.stStationsNummern := stStationsNummern;
Antrieb_Slave.rpRuckzeit        := ppAntriebsInformationenSlave.rpMaxRuckzeit;

// Aufruf Scheibenmessung
Scheibenmessung( stStationsNummern                   := stStationsNummern,
                 ppAntrieb                           := Antrieb,
                 pbpVorstopSensor                    := bpSensorAuslaufVorab,
                 pbpEinlaufSensor                    := bpSensorEinlauf,
                 bpDrehrichtungsumkehrMessung        := bpMessrichtungNegativ,
                 rpMessstrecke                       := ppParameterBaustein.rMessstrecke,
                 ppAntriebsInformationen             := ppAntriebsInformationen,
                 bpAuswahlSensorVorabScheibenmessung := bgFALSE,
                 epGlastyp                           := wpGlastyp,
                 rpFaktorBremswegverlaengern         := 1.6 ) ;
END_FUNCTION_BLOCK

(* ---- Shuttle_Greifer_FB_V01_00_00.fb.st ---- *)
(* METADATA
{
	"v3Meta": {
		"objectGuid": "bb2ac76d-e136-43b9-91b5-1f4b010b201a"
	}
}
*)
FUNCTION_BLOCK Shuttle_Greifer_FB_V01_00_00
VAR_INPUT

  // BOOLEAN
  bpAktivieren                            : BOOL := FALSE; // WICHTIG: Aktivieren des Bausteins (stStationsAufbau.bGreifer)
  bpFreigabe                              : BOOL; // STATUS: Der Greifer ist freigegeben und kann Prozesse abarbeiten
  bpFreigabePneumatik                     : BOOL; // FREIGABE Pneumatik: Greifer-Hub, Greiferzangen, Glasrueckhalter
  bpAutomatikAktiv                        : BOOL;
  bpTeilnehmerErreichbar                  : BOOL;
  bpReset                                 : BOOL;
  bpFahreReferenz                         : BOOL; // BETRIEBSMODUS: Greiferachse referenzieren
  bpCheck                                 : BOOL; // BETRIEBSMODUS: Systemcheck
  bpStartGrundstellungsfahrt              : BOOL; // BETRIEBSMODUS: Grundstellungsfahrt
  bpPositionieren                         : BOOL; // BETRIEBSMODUS: Greifer hinter die Glaskante positionieren (Laenge aus rpGlaslaenge)
  bpStarteVorabPositionierungEintransport : BOOL; // BETRIEBSMODUS: Greifer vor einem Eintransport an die Wandseite stellen
  bpStarteEintransport                    : BOOL; // BETRIEBSMODUS: Scheibe aus dem Faecherwagen auf das Shuttle ziehen
  bpStarteAustransport                    : BOOL; // BETRIEBSMODUS: Scheibe vom Shuttle in den Faecherwagen schieben
  bpSlaveKopplungAktiv                    : BOOL; // STATUS: Glastransport ist auf die Greiferachse gekoppelt
  bpKorrekturfahrtBeendet                 : BOOL; // STATUS: Korrekturfahrt des Glastransports bei uebergrosser Scheibe abgeschlossen
  bpSensorEinlauf                         : BOOL; // STATUS: Einlaufsensor
  bpSensorAuslauf                         : BOOL; // STATUS: Auslaufsensor

  // HANDBETRIEB
  bpHandfahrenPlus                        : BOOL; // Greiferachse in positive Richtung
  bpHandfahrenMinus                       : BOOL; // Greiferachse in negative Richtung
  bpHandGreiferAusfahren                  : BOOL;
  bpHandGreiferEinfahren                  : BOOL;
  bpHandZangeSchliessen                   : BOOL;
  bpHandZangeOeffnen16mm                  : BOOL;
  bpHandZangeOeffnen23mm                  : BOOL;
  bpHandZangeOeffnen29mm                  : BOOL;
  bpHandGlasRueckhalterAusfahren          : BOOL;

  // ENUM
  epGreiferTyp                            : Greifertyp_EN; // AUFTRAGSDATEN: Greiferseite, eGreiferDefault = Seite aus der MK

  // REAL
  rpGlaslaenge                            : REAL; // Scheibenlaenge fuer das Positionieren hinter die Glaskante

  // STRUCT
  pAuftrag                                : Auftragsdaten_ST; // AUFTRAG: Aktuelle Daten zum Auftrag [Laenge, Hoehe, Dicke, Zangenstellung]
  stStationsNummern                       : Station_ST;

  // POINTER
  ppParameterGreifer                      : REFERENCE TO Parameter_Greifer;
  ppAntriebsInformationen                 : REFERENCE TO AntriebsInformationen;

END_VAR
VAR_OUTPUT

  // BOOLEAN
  bpDone                                         : BOOL; // Reset bzw. Referenz abgeschlossen
  bpFehler                                       : BOOL;
  bprtScheibe                                    : BOOL; // Scheibe quittieren
  bpIstInReferenz                                : BOOL;
  bpSicherePosition                              : BOOL; // WICHTIG: Greifer ragt nicht ueber das Shuttle -> Querfahrt erlaubt
  bpGlasRueckhalterEingefahren                   : BOOL; // WICHTIG: Glasrueckhalter eingefahren -> Querfahrt erlaubt
  bpAnforderungSlaveKopplung                     : BOOL; // Anforderung: Glastransport auf die Greiferachse koppeln
  bpKorrekturfahrtAnfordern                      : BOOL; // Anforderung: Glastransport zieht den Rest einer uebergrossen Scheibe auf das Shuttle
  bpKorrekturfahrtRueckwaerts                    : BOOL; // Richtung der Korrekturfahrt: Sensor der Greiferseite frei fahren
  bpAuftragAktiv                                 : BOOL;
  bpVorpositioniertEintransport                  : BOOL; // Greifer steht ausgefahren an der Wandseite fuer den Eintransport
  bpPositionierungAbgeschlossen                  : BOOL;
  bpVorabPositionierungEintransportAbgeschlossen : BOOL;
  bpEintransportAbgeschlossen                    : BOOL;
  bpAustransportAbgeschlossen                    : BOOL;
  bpGrundstellungsfahrtAbgeschlossen             : BOOL;
  bpSystemCheckAbgeschlossen                     : BOOL;

  // WORD
  wpFehlerNr                                     : Fehlerkonstanten_EN;
  wpFehlerKennung                                : WORD; // Zylinder-Kennung bei Zylinderfehlern (cZYLINDER_*), sonst cZYLINDER_KEINE
  awpFehlerInformationen                        : ARRAY[0..25] OF WORD;

  // REAL
  rpWegGlasUebergabeposition                     : REAL; // Weg der Scheibe ueber den Sensor der Greiferseite vor dem Austransport
  rpIstPosition                                  : REAL;

  // ENUM
  epGreiferTypAktiv                              : Greifertyp_EN; // Greiferseite, mit der gearbeitet wird

END_VAR
VAR

  // BOOLEAN
  blErsterZyklus              : BOOL := TRUE;
  blReduzierteGeschwindigkeit : BOOL;
  blUebergrosseScheibe        : BOOL; // Scheibe zu lang, um sie komplett mit dem Greifer zu ziehen
  blSensorSeite               : BOOL; // Sensor der Greiferseite
  blSensorGegenseite          : BOOL; // Sensor der gegenueberliegenden Seite
  blHandAktiv                 : BOOL;
  blZangeSeiteVorhanden       : BOOL; // Greiferzange der aktiven Greiferseite laut MK vorhanden
  blCheckScheibeZiehen        : BOOL; // Systemcheck: Scheibe im Greifer wird auf das Shuttle gezogen (sonst in den Faecherwagen geschoben)
  blCheckNichtQuittieren      : BOOL; // Systemcheck: Greiferzange war offen, die Scheibe wird nicht quittiert
  ablRueckhalterAusfahren     : ARRAY[cZANGE_EINLAUF..cZANGE_AUSLAUF] OF BOOL;

  // INT
  ilZange                     : INT; // Greiferzange der aktiven Seite

  // REAL
  rlRichtung                  : REAL; // +1 Einlaufseite, -1 Auslaufseite: Richtung "auf das Shuttle"
  rlWegBisZumSensor           : REAL;
  rlUebernahmePosition        : REAL;
  rlUebergabePosition         : REAL;
  rlGrundstellungsPosition    : REAL;
  rlGrundstellungGegenseite   : REAL;
  rlGrundstellungEintransport : REAL;
  rlEintransportOffset        : REAL;
  rlPositionUebergrosseScheibe: REAL;
  rlKorrekturOffset           : REAL;
  rlPositionAntriebBeiStart   : REAL;
  rlZielPosition              : REAL;
  rlGlasgewicht               : REAL;

  // ENUM
  elZangeOeffnung             : PneumatikZylinderStatus_EN;

  // STEPS
  steplEintransport                      : Steps_TE;
  steplEintransportMerker                : Steps_TE;
  steplAustransport                      : Steps_TE;
  steplAustransportMerker                : Steps_TE;
  steplPositionieren                     : Steps_TE;
  steplPositionierenMerker               : Steps_TE;
  steplVorabPositionierungEintransport   : Steps_TE;
  steplVorabPositionierungMerker         : Steps_TE;
  steplGrundstellungsfahrt               : Steps_TE;
  steplGrundstellungsfahrtMerker         : Steps_TE;
  steplCheck                             : Steps_TE;
  steplCheckMerker                       : Steps_TE;
  steplReset                             : Steps_TE;
  steplReferenz                          : Steps_TE;
  steplReferenzMerker                    : Steps_TE;

  // TIMER
  tonlAntriebFreigegeben                 : TON; // Endstufe nach "Regler bereit" sicher durchgeschaltet
  tonlMaxWarteAufResetErfolgreich        : TON;
  toflReglerFreigabeErhalten             : TOF; // Reglerfreigabe fuer eine bestimmte Zeit erhalten
  toflSensorSeite                        : TOF; // Entprellen Sensor der Greiferseite
  tonlEndschalterFreifahren              : TON;
  tofHardwareEndschalterFrei             : TOF;
  tonlWarteSchrittEndschalterFreifahren  : TON;
  tonlUeberwachungEintransport           : TON; // Zeitueberwachung der Wartestellen je Schrittkette
  tonlUeberwachungAustransport           : TON;
  tonlUeberwachungPositionieren          : TON;
  tonlUeberwachungVorab                  : TON;
  tonlUeberwachungGrundstellung          : TON;
  tonlUeberwachungCheck                  : TON;
  tonlUeberwachungReferenz               : TON;

  // BAUSTEINE
  Antrieb      : REFERENCE TO Rexroth_ctrlX_Drive_Eckelmann_MC_V01_02_02;
  GreiferHub   : ZylinderPneumatik_FB_V01_00_00; // Greifer aus- / einfahren (ausgefahren = auf Glashoehe)
  Zange        : ARRAY[cZANGE_EINLAUF..cZANGE_AUSLAUF] OF Greiferzange_FB_V01_00_00;

END_VAR
VAR

  // HARDWARE EINGAENGE
  in_bGreiferAusgefahren                 AT %I* : BOOL; // STATUS: Zylinderabfrage Greifer ausgefahren
  in_bGreiferEingefahren                 AT %I* : BOOL; // STATUS: Zylinderabfrage Greifer eingefahren
  in_bGlasRueckhalterEinlaufEingefahren  AT %I* : BOOL; // STATUS: Glasrueckhalter Einlaufseite eingefahren
  in_bGlasRueckhalterAuslaufEingefahren  AT %I* : BOOL; // STATUS: Glasrueckhalter Auslaufseite eingefahren

  // HARDWARE AUSGAENGE
  out_bGreiferAusfahren                  AT %Q* : BOOL; // Impuls Zylinder Greifer ausfahren
  out_bGreiferEinfahren                  AT %Q* : BOOL; // Impuls Zylinder Greifer einfahren
  out_bGlasRueckhalterEinlaufAusfahren   AT %Q* : BOOL; // Federrueckstellventil Glasrueckhalter Einlaufseite: TRUE = ausgefahren
  out_bGlasRueckhalterAuslaufAusfahren   AT %Q* : BOOL; // Federrueckstellventil Glasrueckhalter Auslaufseite: TRUE = ausgefahren

END_VAR
VAR CONSTANT

  // INT
  cZANGE_EINLAUF      : INT := 1;
  cZANGE_AUSLAUF      : INT := 2;

  // REAL
  cTOLERANZ_POSITION  : REAL := 2.5; // [mm] Zielposition erreicht

  // TIME
  cZEIT_SENSOR_ENTPRELLEN : TIME := T#50MS;

END_VAR
(* Anmerkung:
   - Greifer im Shuttle: eigene Greiferachse, Greifer aus-/einfahren, Greiferzange und Glasrueckhalter je Seite
     optional (Parameter_Greifer.bZange...Vorhanden / bGlasRueckhalter...Vorhanden)
   - Ablaeufe ueber eine Greiferseite ohne Greiferzange werden mit Meldung abgelehnt
   - Eintransport: Scheibe im Faecherwagen greifen und auf das Shuttle ziehen, der Glastransport ist dabei
     auf die Greiferachse gekoppelt (Slave)
   - Austransport: Scheibe greifen und in den Faecherwagen schieben
*)
//-------------------------------------------------------------------------------------------------
// BAUSTEIN: DEAKTIVIERUNG
//-------------------------------------------------------------------------------------------------
(* Hinweis:
   - Ein deaktivierter Greifer meldet kein Done und keine Status-Freigaben; der Aufrufer verknuepft
     mit der Aktivierung aus der MK (z.B. Greifer.bpSicherePosition OR NOT stStationsAufbau.bGreifer[wWand])
*)
IF ( NOT bpAktivieren ) THEN

  out_bGreiferAusfahren                := FALSE;
  out_bGreiferEinfahren                := FALSE;
  out_bGlasRueckhalterEinlaufAusfahren := FALSE;
  out_bGlasRueckhalterAuslaufAusfahren := FALSE;

  ablRueckhalterAusfahren[cZANGE_EINLAUF] := FALSE;
  ablRueckhalterAusfahren[cZANGE_AUSLAUF] := FALSE;

  GreiferHub();
  Zange[cZANGE_EINLAUF]();
  Zange[cZANGE_AUSLAUF]();

  bpDone                                         := FALSE;
  bpFehler                                       := FALSE;
  wpFehlerNr                                     := cMELDUNG_NULL;
  wpFehlerKennung                                := cZYLINDER_KEINE;
  bprtScheibe                                    := FALSE;
  bpIstInReferenz                                := FALSE;
  bpSicherePosition                              := FALSE;
  bpGlasRueckhalterEingefahren                   := FALSE;
  bpAnforderungSlaveKopplung                     := FALSE;
  bpKorrekturfahrtAnfordern                      := FALSE;
  bpAuftragAktiv                                 := FALSE;
  bpVorpositioniertEintransport                  := FALSE;
  bpPositionierungAbgeschlossen                  := FALSE;
  bpVorabPositionierungEintransportAbgeschlossen := FALSE;
  bpEintransportAbgeschlossen                    := FALSE;
  bpAustransportAbgeschlossen                    := FALSE;
  bpGrundstellungsfahrtAbgeschlossen             := FALSE;
  bpSystemCheckAbgeschlossen                     := FALSE;

  RETURN;

END_IF

//-------------------------------------------------------------------------------------------------
// BAUSTEIN: INITIALISIERUNG
//-------------------------------------------------------------------------------------------------
IF ( blErsterZyklus ) THEN

  IF ( __ISVALIDREF(ppAntriebsInformationen) AND __ISVALIDREF(ppParameterGreifer) ) THEN

    blErsterZyklus := FALSE;

    Antrieb REF= pgAntriebe[ppAntriebsInformationen.wAchsID];

    (* Hinweis:
       - Initialisierung Antriebsinformationen
    *)
    Antrieb.ppAntriebsInformationen REF= ppAntriebsInformationen;
    Antrieb.rpZielPosition    := Antrieb.rpIstPosition;
    Antrieb.rpGeschwindigkeit := ppAntriebsInformationen.rpMaxGeschwindigkeit;
    Antrieb.rpBeschleunigung  := ppAntriebsInformationen.rpMaxBeschleunigung;
    Antrieb.rpVerzoegerung    := ppAntriebsInformationen.rpMaxVerzoegerung;
    Antrieb.rpRuckzeit        := ppAntriebsInformationen.rpMaxRuckzeit;

    (* Hinweis:
       - Pneumatik: Greifer mit Endlagenabfragen, Greiferzangen laut MK
       - Eine nicht vorhandene Greiferzange ist deaktiviert (keine Ausgaenge, kein Done, kein Fehler)
    *)
    GreiferHub.bpAktivieren                  := TRUE;
    GreiferHub.bpAbfrageAusgefahrenVorhanden := TRUE;
    GreiferHub.bpAbfrageEingefahrenVorhanden := TRUE;

    Zange[cZANGE_EINLAUF].bpAktivieren := ppParameterGreifer.bZangeEinlaufVorhanden;
    Zange[cZANGE_AUSLAUF].bpAktivieren := ppParameterGreifer.bZangeAuslaufVorhanden;

  ELSE
    RETURN;
  END_IF

END_IF

//-------------------------------------------------------------------------------------------------
// BAUSTEIN: GREIFERSEITE
//-------------------------------------------------------------------------------------------------
(* Hinweis:
   - Seite aus dem Auftrag, sonst aus der MK
   - rlRichtung: Richtung der Greiferachse "auf das Shuttle" (Einlaufseite positiv, Auslaufseite negativ)
*)
IF ( epGreiferTyp <> eGreiferDefault ) THEN
  epGreiferTypAktiv := epGreiferTyp;
ELSE
  epGreiferTypAktiv := ppParameterGreifer.eGreiferTyp;
END_IF

IF ( epGreiferTypAktiv = eGreiferAuslaufseite ) THEN
  ilZange                      := cZANGE_AUSLAUF;
  rlRichtung                   := -1.0;
  rlWegBisZumSensor            := ppParameterGreifer.rWegBisZumAuslaufsensor;
  rlUebernahmePosition         := ppParameterGreifer.rUebernahmePosition_Auslauf;
  rlUebergabePosition          := ppParameterGreifer.rUebergabePosition_Auslauf;
  rlGrundstellungsPosition     := ppParameterGreifer.rGrundstellungsPosition_Auslauf;
  rlGrundstellungGegenseite    := ppParameterGreifer.rGrundstellungsPosition_Einlauf;
  rlGrundstellungEintransport  := ppParameterGreifer.rGrundstellungsPosition_AuslaufEintransport;
  rlPositionUebergrosseScheibe := ppParameterGreifer.rPositionUebergrosseScheibe_Auslauf;
  rlKorrekturOffset            := ppParameterGreifer.rKorrekturOffset_Auslauf;
  blSensorSeite                := bpSensorAuslauf;
  blSensorGegenseite           := bpSensorEinlauf;
  IF ( pAuftrag.bLetzteScheibe ) THEN
    rlEintransportOffset := ppParameterGreifer.rGlasEintransportOffset_Auslauf;
  ELSE
    rlEintransportOffset := ppParameterGreifer.rGlasEintransportOffset_AuslaufSammeln;
  END_IF
ELSE
  ilZange                      := cZANGE_EINLAUF;
  rlRichtung                   := 1.0;
  rlWegBisZumSensor            := ppParameterGreifer.rWegBisZumEinlaufsensor;
  rlUebernahmePosition         := ppParameterGreifer.rUebernahmePosition_Einlauf;
  rlUebergabePosition          := ppParameterGreifer.rUebergabePosition_Einlauf;
  rlGrundstellungsPosition     := ppParameterGreifer.rGrundstellungsPosition_Einlauf;
  rlGrundstellungGegenseite    := ppParameterGreifer.rGrundstellungsPosition_Auslauf;
  rlGrundstellungEintransport  := ppParameterGreifer.rGrundstellungsPosition_EinlaufEintransport;
  rlPositionUebergrosseScheibe := ppParameterGreifer.rPositionUebergrosseScheibe_Einlauf;
  rlKorrekturOffset            := ppParameterGreifer.rKorrekturOffset_Einlauf;
  blSensorSeite                := bpSensorEinlauf;
  blSensorGegenseite           := bpSensorAuslauf;
  IF ( pAuftrag.bLetzteScheibe ) THEN
    rlEintransportOffset := ppParameterGreifer.rGlasEintransportOffset_Einlauf;
  ELSE
    rlEintransportOffset := ppParameterGreifer.rGlasEintransportOffset_EinlaufSammeln;
  END_IF
END_IF

bpKorrekturfahrtRueckwaerts := ( epGreiferTypAktiv = eGreiferAuslaufseite );

(* Hinweis:
   - Ohne Greiferzange auf der aktiven Seite lehnen Ein-/Austransport, Positionieren, Vorabpositionierung
     und Systemcheck mit cMELDUNG_AUFTRAGSDATEN_SHUTTLE_GREIFER_AUFTRAGSTYP_UNGUELTIG ab
*)
blZangeSeiteVorhanden :=    ( ( ilZange = cZANGE_EINLAUF ) AND ppParameterGreifer.bZangeEinlaufVorhanden )
                         OR ( ( ilZange = cZANGE_AUSLAUF ) AND ppParameterGreifer.bZangeAuslaufVorhanden );

(* Hinweis:
   - Uebergrosse Scheibe: der Greifer zieht nur bis rPositionUebergrosseScheibe, den Rest zieht der Glastransport
   - Oeffnung der Greiferzange aus dem Auftrag, ohne Vorgabe maximal geoeffnet
*)
blUebergrosseScheibe := ( pAuftrag.rAuftragsLaenge >= ppParameterGreifer.rLaengeUebergroesseScheibe )
                        AND ( ppParameterGreifer.rLaengeUebergroesseScheibe > 0.0 );

IF ( blUebergrosseScheibe ) THEN
  rpWegGlasUebergabeposition := ppParameterGreifer.rWegGlasUebergabepositionLang;
ELSE
  rpWegGlasUebergabeposition := ppParameterGreifer.rWegGlasUebergabeposition;
END_IF

IF (    ( pAuftrag.stAuftragsOptionen.eGreiferZangeStellung = eZylinderStellung16mm )
     OR ( pAuftrag.stAuftragsOptionen.eGreiferZangeStellung = eZylinderStellung23mm )
     OR ( pAuftrag.stAuftragsOptionen.eGreiferZangeStellung = eZylinderStellung29mm ) )
THEN
  elZangeOeffnung := pAuftrag.stAuftragsOptionen.eGreiferZangeStellung;
ELSE
  elZangeOeffnung := eZylinderStellung29mm;
END_IF

//-------------------------------------------------------------------------------------------------
// BAUSTEIN: TIMER, EINSTELLUNGEN, ETC.
//-------------------------------------------------------------------------------------------------
(* Hinweis:
   - Die Endstufe des Umrichters ist bei "bpReglerBereit" noch nicht sicher durchgeschaltet
*)
tonlAntriebFreigegeben( IN := Antrieb.bpReglerBereit, PT := T#200MS );

tonlMaxWarteAufResetErfolgreich( IN := bpReset, PT := tgMaxWartezeitReset - T#1S );

toflSensorSeite( IN := blSensorSeite, PT := cZEIT_SENSOR_ENTPRELLEN );

//-------------------------------------------------------------------------------------------------
// BAUSTEIN: AKTIONEN
//-------------------------------------------------------------------------------------------------
SystemCheck();

Positionieren();
VorabPositionierungEintransport();
Eintransport();
Austransport();
Grundstellung();

Reset();
Referenz();
Handfunktionen();
Meldungen();

//-------------------------------------------------------------------------------------------------
// BAUSTEIN: SICHERHEIT UND STATUS
//-------------------------------------------------------------------------------------------------
(* Hinweis:
   - Greifer ragt nicht ueber die Aussenkanten des Shuttles
   - Glasrueckhalter eingefahren (ein nicht vorhandener Glasrueckhalter gilt als eingefahren)
*)
bpSicherePosition := (     Antrieb.bpIstReferenziert
                       AND ( Antrieb.rpIstPosition >= ppParameterGreifer.rSicherPositionMinimal )
                       AND ( Antrieb.rpIstPosition <= ppParameterGreifer.rSicherPositionMaximal ) );

bpGlasRueckhalterEingefahren :=     ( in_bGlasRueckhalterEinlaufEingefahren OR NOT ppParameterGreifer.bGlasRueckhalterEinlaufVorhanden )
                                AND ( in_bGlasRueckhalterAuslaufEingefahren OR NOT ppParameterGreifer.bGlasRueckhalterAuslaufVorhanden );

bpIstInReferenz := Antrieb.bpIstReferenziert;
rpIstPosition   := Antrieb.rpIstPosition;

bpAuftragAktiv :=    ( bpStarteEintransport AND ( steplEintransport > STEP_0_E ) )
                  OR ( bpStarteAustransport AND ( steplAustransport > STEP_0_E ) )
                  OR ( bpPositionieren AND ( steplPositionieren > STEP_0_E ) )
                  OR ( bpStarteVorabPositionierungEintransport AND ( steplVorabPositionierungEintransport > STEP_0_E ) )
                  OR ( bpStartGrundstellungsfahrt AND ( steplGrundstellungsfahrt > STEP_0_E ) );

//-------------------------------------------------------------------------------------------------
// BAUSTEIN: FREIGABEN UND AUFRUFE
//-------------------------------------------------------------------------------------------------
toflReglerFreigabeErhalten( IN := (    bpHandfahrenPlus
                                    OR bpHandfahrenMinus
                                    OR bpFahreReferenz
                                    OR bpCheck
                                    OR bpStarteEintransport
                                    OR bpStarteAustransport
                                    OR bpPositionieren
                                    OR bpStarteVorabPositionierungEintransport
                                    OR bpStartGrundstellungsfahrt ),
                            PT := ppParameterGreifer.tZeitAntriebsfreigabeErhalten );

// Aufruf Antrieb (der Antrieb selbst wird zentral im Programm Antriebe aufgerufen)
Antrieb.bpFreigabe        := bpFreigabe AND toflReglerFreigabeErhalten.Q;
Antrieb.stStationsNummern := stStationsNummern;
Antrieb.rpRuckzeit        := ppAntriebsInformationen.rpMaxRuckzeit;

// Aufruf Pneumatik
GreiferHub( bpFreigabe                    := bpFreigabePneumatik,
            in_bStatusZylinderAusgefahren := in_bGreiferAusgefahren,
            in_bStatusZylinderEingefahren := in_bGreiferEingefahren );

Zange[cZANGE_EINLAUF]( bpFreigabe := bpFreigabePneumatik, bpZylinderAbfragenVorhanden := ppParameterGreifer.bZangeAbfragenVorhanden, tpBewegungszeit := ppParameterGreifer.tZangeBewegungszeit );
Zange[cZANGE_AUSLAUF]( bpFreigabe := bpFreigabePneumatik, bpZylinderAbfragenVorhanden := ppParameterGreifer.bZangeAbfragenVorhanden, tpBewegungszeit := ppParameterGreifer.tZangeBewegungszeit );

//-------------------------------------------------------------------------------------------------
// BAUSTEIN: AUSGAENGE
//-------------------------------------------------------------------------------------------------
out_bGreiferAusfahren := GreiferHub.out_bZylinderAusfahren;
out_bGreiferEinfahren := GreiferHub.out_bZylinderEinfahren;

out_bGlasRueckhalterEinlaufAusfahren := ablRueckhalterAusfahren[cZANGE_EINLAUF] AND ppParameterGreifer.bGlasRueckhalterEinlaufVorhanden AND bpFreigabePneumatik;
out_bGlasRueckhalterAuslaufAusfahren := ablRueckhalterAusfahren[cZANGE_AUSLAUF] AND ppParameterGreifer.bGlasRueckhalterAuslaufVorhanden AND bpFreigabePneumatik;
END_FUNCTION_BLOCK

(* ---- Shuttle_Kippen_V01_00_00.fb.st ---- *)
(* METADATA
{
	"v3Meta": {
		"objectGuid": "188879d4-0bd4-40ef-906f-fea4dde7d858"
	}
}
*)
FUNCTION_BLOCK Shuttle_Kippen_V01_00_00
VAR_INPUT

  // BOOL
  bpSensorEinlauf                  : BOOL;
  bpSensorAuslauf                  : BOOL;
  bpAktivieren                     : BOOL;
  bpPositionieren                  : BOOL;
  bpReset                          : BOOL;
  bpReferenz                       : BOOL;
  bpBetriebsartHand                : BOOL;
  bpFreigabe                       : BOOL;
  bpLangsamKippen                  : BOOL;
  bpTeilnehmerErreichbar           : BOOL;
  bpKippenSchuetz                  : BOOL;

  // STRUCT
  stStationsNummern      : Station_ST;
  epZielPosition         : Kippen_EN;

  // POINTER
  ppParameterBaustein     : REFERENCE TO Parameter_Kippen;
  ppAntriebsInformationen : REFERENCE TO AntriebsInformationen;

END_VAR
VAR_OUTPUT

  // BOOL
  bpDone                 : BOOL;
  bpFehler               : BOOL;
  bpInReferenz           : BOOL;

  // WORD
  wpFehlerNr             : Fehlerkonstanten_EN;

  // REAL
  rpAktuelleKippPosition : REAL;
  rpOutGeschwindigkeit   : REAL;

  // ENUM
  epKippStatus           : Kippen_EN;

END_VAR
VAR

  // BOOL
  blErsterZyklus                : BOOL := TRUE;
  blSensorEinlauf               : BOOL;
  blSensorAuslauf               : BOOL;
  bpStartAufkippen              : BOOL;
  bpStartAbkippen               : BOOL;

  // TIMER
  tonlMaxWarteAufResetErfolgreich       : TON;
  tonlAntriebNichtFreigegeben           : TON; // Ueberwachung: Antrieb nicht betriebsbereit
  tonlEndschalterFreifahren             : TON;
  tonlWarteSchrittEndschalterFreifahren : TON;
  tofHardwareEndschalterFrei            : TOF;
  toflReglerFreigabeErhalten            : TOF;
  tonlSensorEinlauf                     : TON;
  tonlSensorAuslauf                     : TON;
  toflReset                             : TOF;
  tonlTeilnehmerErreichbar              : TON;
  tonlMaxWarteZeit                      : TON;
  toflMotorstarterOK                    : TOF;
  toflMotorSicherungOK                  : TOF;

  // STEPS
  steplPositionieren : Steps_TE;
  steplReferenz      : Steps_TE;
  steplReset         : Steps_TE;
  steplKippenSchuetz : Steps_TE; // Mit Schütz Kippen

  // Antrieb
  Antrieb : REFERENCE TO Rexroth_ctrlX_Drive_Eckelmann_MC_V01_02_02;

END_VAR
VAR

  // HARDWARE EINGAENGE
  in_bMotorschutzschalter_OK           AT %I* : BOOL;
  in_bLeitungsschutzschalterBremseOK   AT %I* : BOOL;
  in_bMotorstarter_OK           : BOOL;
  in_bSensorNicht90Grad         : BOOL;
  in_bSensorNicht84Grad         : BOOL;

  // HARDWARE AUSGAENGE
  out_bKippenAbSetzen           : BOOL;
  out_bKippenAufSetzen          : BOOL;
  out_bBremseLoesen             : BOOL;
  out_bReset                    : BOOL;

END_VAR
//-------------------------------------------------------------------------------------------------
// INITIALISIERUNG
//-------------------------------------------------------------------------------------------------
IF ( blErsterZyklus ) THEN

  IF ( __ISVALIDREF(ppAntriebsInformationen) ) THEN

    blErsterZyklus := FALSE;

    Antrieb REF= pgAntriebe[ppAntriebsInformationen.wAchsID];

    (* Hinweis:
       - Initialisierung Antriebsinformationen
    *)
    Antrieb.ppAntriebsInformationen REF= ppAntriebsInformationen;

    (* Hinweis:
       - Für die Zielpunktkontrolle muss im ersten Zyklus die Zielposition initialisiert werden
    *)
    Antrieb.rpZielPosition := Antrieb.rpIstPosition;

    (* Hinweis:
       - Antriebswerte vorinitialisieren
    *)
    Antrieb.rpGeschwindigkeit := ppAntriebsInformationen.rpMaxGeschwindigkeit;
    Antrieb.rpBeschleunigung  := ppAntriebsInformationen.rpMaxBeschleunigung;
    Antrieb.rpVerzoegerung    := ppAntriebsInformationen.rpMaxVerzoegerung;
    Antrieb.rpRuckzeit        := ppAntriebsInformationen.rpMaxRuckzeit;

    tonlTeilnehmerErreichbar(IN := FALSE);
    tonlMaxWarteZeit(IN := FALSE);

  ELSE
    RETURN;
  END_IF

END_IF

// Endschalter zyklisch an den Antrieb geben: 84 Grad = Min, 90 Grad = Max (Oeffner, wirkt nur bei Endschalterquelle SPS)
Antrieb.bpEndschalterMaxExtern := in_bSensorNicht90Grad;
Antrieb.bpEndschalterMinExtern := in_bSensorNicht84Grad;

//-------------------------------------------------------------------------------------------------
// DEAKTIVIEREN
//-------------------------------------------------------------------------------------------------

IF ( NOT bpAktivieren ) THEN
  bpDone     := TRUE;
  bpFehler   := FALSE;
  wpFehlerNr := cMELDUNG_NULL;

  IF ( bpPositionieren AND ( epZielPosition = eKippen_Position_0Grad ) ) THEN
    epKippStatus := eKippen_Position_0Grad;
  ELSIF ( bpPositionieren AND ( epZielPosition = eKippen_Position_84Grad ) ) THEN
    epKippStatus := eKippen_Position_84Grad;
  ELSIF ( bpPositionieren AND ( epZielPosition = eKippen_Position_88_5Grad ) ) THEN
    epKippStatus := eKippen_Position_88_5Grad;
  ELSIF ( bpPositionieren AND ( epZielPosition = eKippen_Position_90Grad ) ) THEN
    epKippStatus := eKippen_Position_90Grad;
  ELSIF ( bpPositionieren AND ( epZielPosition = eKippen_Position_96Grad ) ) THEN
    epKippStatus := eKippen_Position_96Grad;
  ELSE
    epKippStatus := eKippen_Default;
  END_IF

  RETURN;

END_IF

//-------------------------------------------------------------------------------------------------
// TIMER
//-------------------------------------------------------------------------------------------------
// Reset- Ueberwachung
tonlMaxWarteAufResetErfolgreich(IN := bpReset, pt := tgMaxWartezeitReset-T#1S);
tonlSensorEinlauf( IN := bpSensorEinlauf , pt := T#200MS );
tonlSensorAuslauf( IN := bpSensorAuslauf , pt := T#200MS );
blSensorEinlauf := tonlSensorEinlauf.Q;
blSensorAuslauf := tonlSensorAuslauf.Q;

tonlTeilnehmerErreichbar( IN := bpTeilnehmerErreichbar, PT := T#5S );
tonlMaxWarteZeit(IN:=(    ( bpStartAbKippen AND out_bKippenAbSetzen )
                       OR ( bpStartAufKippen AND out_bKippenAufSetzen ) ),
                  PT:= ppParameterBaustein.tZeitlicheUeberwachungKippen );

//-------------------------------------------------------------------------------------------------
// AKTIONEN
//-------------------------------------------------------------------------------------------------
Meldungen();
Ausgaenge();
Reset();

IF ( bpKippenSchuetz ) THEN
  // Bremse lösen
  out_bBremseLoesen := out_bKippenAbSetzen OR out_bKippenAufSetzen OR bgVISUKippenBremseLoesen[stStationsNummern.NummerSPS];

  // Reset Motorstarter
  toflReset( IN := bpReset, PT := T#3S );
  out_bReset := toflReset.Q;

  Kippen_Schuetz();

ELSE
  Positionieren();
  Referenz();

  IF ( NOT bpKippenSchuetz ) THEN
    // Antriebsfreigabe:
    toflReglerFreigabeErhalten( IN := (   bpPositionieren
                                        OR bpReferenz ),
                                PT := ppParameterBaustein.tZeitAntriebsfreigabeErhalten );

    // Aufruf
    Antrieb.bpFreigabe        := bpFreigabe AND toflReglerFreigabeErhalten.Q;
    Antrieb.rpRuckzeit        := ppAntriebsInformationen.rpMaxRuckzeit;
    Antrieb.stStationsNummern := stStationsNummern;

  END_IF

END_IF
END_FUNCTION_BLOCK

(* ---- Wandverstellung_MultiZylinder_FB_V01_00_00.fb.st ---- *)
(* METADATA
{
	"v3Meta": {
		"objectGuid": "57ebb36f-f22e-4632-9b59-8f205a70f04c"
	}
}
*)
FUNCTION_BLOCK Wandverstellung_MultiZylinder_FB_V01_00_00
VAR_INPUT

  // BOOLEAN
  bpReset                     : BOOL;
  bpAktivieren                : BOOL;
  bpFreigabe                  : BOOL; // FREIGABE Pneumatik: ohne Freigabe Ventile aus, Bewegung pausiert (Startbefehl bleibt erhalten)
  bpStartZylinderBewegung     : BOOL; // BETRIEBTYP: Zylinder wird ausgefahren
  bpZylinderAbfragenVorhanden : BOOL := FALSE; // Hinweis: Manche Zylinder haben keine Abfragen

  // TIME
  tpBewegungszeit             : TIME := T#1S; // Bewegungszeit je Richtung ohne Abfragen

  // ENUM
  epSollZylinderStellung  : PneumatikZylinderStatus_EN;

END_VAR

VAR_OUTPUT

  // BOOLEAN
  bpFehler                       : BOOL;
  bpDone                         : BOOL;

  // WORD
  wpFehlerNr       : Fehlerkonstanten_EN;

  // ENUM
  epStatusZylinderStellung : PneumatikZylinderStatus_EN;

END_VAR

VAR

  // STEPS
  steplZylinderStellung   : Steps_TE;

  // TIMER
  tonlStellung13mm               : TON; // EINSCHALTVERZOEGERUNG: Warten bis der Zylinder eingefahren wurde. Sonst wird ein Fehlerausgegeben
  tonlStellung23mm               : TON; // EINSCHALTVERZOEGERUNG: Warten bis der Zylinder ausgefahren wurde. Sonst wird ein Fehlerausgegeben
  tonlStellung29mm               : TON; // EINSCHALTVERZOEGERUNG: Warten bis der Zylinder eingefahren wurde. Sonst wird ein Fehlerausgegeben
  tonlWartezeitZylinderStellung  : TON; // EINSCHALTVERZOEGERUNG: wenn keine Abfragen verbaut sind, pauschal die Schaltung der Ventile zurücksetzen

END_VAR

VAR

  // HARDWAREEINGAENGE
  in_bStatusZylinder_1_Ausgefahren     AT %I* : BOOL; // STATUS: Zylinderabfrage [Ausgefahren]
  in_bStatusZylinder_2_Ausgefahren     AT %I* : BOOL; // STATUS: Zylinderabfrage [Ausgefahren]
  in_bStatusZylinder_Alle_Eingefahren  AT %I* : BOOL; // STATUS: Zylinderabfrage [Eingefahren]

  // HARDWAREAUSGAENGE
  out_bZylinder_1_Einfahren    AT %Q* : BOOL; // Impuls Zylinder: x mm Hub
  out_bZylinder_2_Einfahren    AT %Q* : BOOL; // Impuls Zylinder: X mm Hub
  out_bZylinder_1_Ausfahren    AT %Q* : BOOL; // Impuls Zylinder: x mm Hub
  out_bZylinder_2_Ausfahren    AT %Q* : BOOL; // Impuls Zylinder: x mm Hub

END_VAR
//-------------------------------------------------------------------------------------------------
// BAUSTEIN: RESET / DEAKTIVIERT
//-------------------------------------------------------------------------------------------------
(* Hinweis:
   - Reset oder deaktiviert: Ausgaenge aus, Kette und Timer zuruecksetzen, Done und Fehler loeschen
   - Der Baustein setzt bpReset selbst zurueck, der Aufrufer wartet nicht auf Done
   - Ein deaktivierter Baustein meldet kein Done; der Aufrufer verknuepft das Warten auf Done
     mit der Aktivierung aus der MK (z.B. Wandverstellung.bpDone OR NOT stStationsAufbau.bX)
*)
IF ( bpReset OR NOT bpAktivieren ) THEN

  out_bZylinder_1_Einfahren := FALSE;
  out_bZylinder_2_Einfahren := FALSE;
  out_bZylinder_1_Ausfahren := FALSE;
  out_bZylinder_2_Ausfahren := FALSE;

  bpStartZylinderBewegung := FALSE;

  steplZylinderStellung := STEP_0_E;

  tonlStellung13mm( IN := FALSE );
  tonlStellung23mm( IN := FALSE );
  tonlStellung29mm( IN := FALSE );
  tonlWartezeitZylinderStellung( IN := FALSE );

  bpDone     := FALSE;
  bpFehler   := FALSE;
  wpFehlerNr := cMELDUNG_NULL;

  bpReset := FALSE;

  RETURN;

END_IF

//-------------------------------------------------------------------------------------------------
// BAUSTEIN: AKTIONEN
//-------------------------------------------------------------------------------------------------
(* Hinweis Freigabe Pneumatik:
   - Ohne Freigabe: Ventile aus, Kette und Ueberwachungszeiten zuruecksetzen (kein Timeout-Fehler)
   - Der Startbefehl bleibt erhalten: kommt die Freigabe zurueck, wird die Bewegung neu gestartet
*)
IF NOT bpFreigabe THEN
  out_bZylinder_1_Einfahren := FALSE;
  out_bZylinder_2_Einfahren := FALSE;
  out_bZylinder_1_Ausfahren := FALSE;
  out_bZylinder_2_Ausfahren := FALSE;
  steplZylinderStellung := STEP_0_E;
  tonlStellung13mm( IN := FALSE );
  tonlStellung23mm( IN := FALSE );
  tonlStellung29mm( IN := FALSE );
  tonlWartezeitZylinderStellung( IN := FALSE );
  bpDone := FALSE;
ELSE
  ZylinderBewegung();
END_IF

//-------------------------------------------------------------------------------------------------
// STATUS DER ZYLINDER
//-------------------------------------------------------------------------------------------------
(* Hinweis:
   - Status aus der Sensorik, wenn Abfragen vorhanden sind
   - Ohne Abfragen bleibt der Status, den die Schrittkette nach der Bewegungszeit setzt
*)
IF ( bpZylinderAbfragenVorhanden ) THEN

  // Stellung 29mm
  IF (     in_bStatusZylinder_1_Ausgefahren
       AND in_bStatusZylinder_2_Ausgefahren )
  THEN
    epStatusZylinderStellung := eZylinderStellung29mm;

  // Stellung 23mm
  ELSIF (     in_bStatusZylinder_1_Ausgefahren
          AND NOT in_bStatusZylinder_2_Ausgefahren )
  THEN
    epStatusZylinderStellung := eZylinderStellung23mm;

  // Stellung 13mm
  ELSIF (     in_bStatusZylinder_Alle_Eingefahren
          AND NOT in_bStatusZylinder_1_Ausgefahren
          AND NOT in_bStatusZylinder_2_Ausgefahren )
  THEN
    epStatusZylinderStellung := eZylinderStellung16mm;

  ELSE
    epStatusZylinderStellung := eZylinderUndefiniert;

  END_IF

END_IF
END_FUNCTION_BLOCK

(* ---- Wandverstellung_Pneumatik_FB_V01_00_00.fb.st ---- *)
(* METADATA
{
	"v3Meta": {
		"objectGuid": "3c575514-d133-4a53-b99b-31124f37ab50"
	}
}
*)
FUNCTION_BLOCK Wandverstellung_Pneumatik_FB_V01_00_00
VAR_INPUT

  // BOOLEAN
  bpWandverstellungOeffnen    : BOOL;
  bpWandverstellungSchliessen : BOOL;
  bpReset                     : BOOL;
  bpAktivieren                : BOOL;
  bpFreigabe                  : BOOL; // FREIGABE Pneumatik: ohne Freigabe Ventile aus, Bewegung pausiert (Startbefehl bleibt erhalten)

  // OPTIONEN
  bpAbfrageGeoeffnetVorhanden   : BOOL := TRUE;   // Endlagensensoren geoeffnet vorhanden, sonst gilt die Endlage nach tpBewegungszeit
  bpAbfrageGeschlossenVorhanden : BOOL := TRUE;   // Endlagensensoren geschlossen vorhanden, sonst gilt die Endlage nach tpBewegungszeit
  tpBewegungszeit               : TIME := T#800MS; // Bewegungszeit je Richtung ohne Endlagensensor

END_VAR
VAR_OUTPUT

  // BOOLEAN
  bpDone    : BOOL;
  bpFehler  : BOOL;

  // WORD
  wpFehlerNr  : Fehlerkonstanten_EN;

END_VAR
VAR

  // STEPS
  steplWandverstellungOeffnen    : Steps_TE;
  steplWandverstellungSchliessen : Steps_TE;

  // TIMER
  tonlEingefahrenWandEinlaufseite  : TON; // EINSCHALTVERZOEGERUNG: Warten bis der Zylinder verfahren wurde. Sonst wird ein Fehlerausgegeben
  tonlAusgefahrenWandEinlaufseite  : TON; // EINSCHALTVERZOEGERUNG: Warten bis der Zylinder verfahren wurde. Sonst wird ein Fehlerausgegeben
  tonlEingefahrenWandAuslaufseite  : TON; // EINSCHALTVERZOEGERUNG: Warten bis der Zylinder verfahren wurde. Sonst wird ein Fehlerausgegeben
  tonlAusgefahrenWandAuslaufseite  : TON; // EINSCHALTVERZOEGERUNG: Warten bis der Zylinder verfahren wurde. Sonst wird ein Fehlerausgegeben
  tonlBewegungszeitOeffnen         : TON; // Bewegungszeit ohne Endlagensensor geoeffnet
  tonlBewegungszeitSchliessen      : TON; // Bewegungszeit ohne Endlagensensor geschlossen

END_VAR
VAR

  // HARDWARE EINGAENGE
  in_bWandEinlaufseiteGeoeffnet    AT %I* : BOOL; // STATUS: Sensor meldet geöffnet
  in_bWandEinlaufseiteGeschlossen  AT %I* : BOOL; // STATUS: Sensor meldet geschlossen
  in_bWandAuslaufseiteGeoeffnet    AT %I* : BOOL; // STATUS: Sensor meldet geöffnet
  in_bWandAuslaufseiteGeschlossen  AT %I* : BOOL; // STATUS: Sensor meldet geschlossen

  // HARDWARE AUSGAENGE
  out_bWandverstellungOeffnen      AT %Q* : BOOL; // AKTION: Verstellen der Wandoeffnung -> Maximal Geoeffnet
  out_bWandverstellungSchliessen   AT %Q* : BOOL; // AKTION: Verstellen der Wandoeffnung -> Minimal Geoeffnet

END_VAR
//-------------------------------------------------------------------------------------------------
// BAUSTEIN: RESET / DEAKTIVIERT
//-------------------------------------------------------------------------------------------------
(* Hinweis:
   - Reset oder deaktiviert: Ausgaenge aus, Ketten und Timer zuruecksetzen, Done und Fehler loeschen
   - Der Baustein setzt bpReset selbst zurueck, der Aufrufer wartet nicht auf Done
   - Ein deaktivierter Baustein meldet kein Done; der Aufrufer verknuepft das Warten auf Done
     mit der Aktivierung aus der MK (z.B. Wandverstellung.bpDone OR NOT stStationsAufbau.bX)
*)
IF ( bpReset OR NOT bpAktivieren ) THEN

  out_bWandverstellungOeffnen    := FALSE;
  out_bWandverstellungSchliessen := FALSE;

  bpWandverstellungOeffnen    := FALSE;
  bpWandverstellungSchliessen := FALSE;

  steplWandverstellungOeffnen    := STEP_0_E;
  steplWandverstellungSchliessen := STEP_0_E;

  tonlEingefahrenWandEinlaufseite( IN := FALSE );
  tonlAusgefahrenWandEinlaufseite( IN := FALSE );
  tonlEingefahrenWandAuslaufseite( IN := FALSE );
  tonlAusgefahrenWandAuslaufseite( IN := FALSE );
  tonlBewegungszeitOeffnen( IN := FALSE );
  tonlBewegungszeitSchliessen( IN := FALSE );

  wpFehlerNr := cMELDUNG_NULL;
  bpFehler   := FALSE;
  bpDone     := FALSE;

  bpReset := FALSE;

  RETURN;

END_IF

//-------------------------------------------------------------------------------------------------
// BAUSTEIN: AKTIONEN
//-------------------------------------------------------------------------------------------------
(* Hinweis Freigabe Pneumatik:
   - Ohne Freigabe: Ventile aus, Ketten und Ueberwachungszeiten zuruecksetzen (kein Timeout-Fehler)
   - Der Startbefehl bleibt erhalten: kommt die Freigabe zurueck, wird die Bewegung neu gestartet
*)
IF NOT bpFreigabe THEN
  out_bWandverstellungOeffnen    := FALSE;
  out_bWandverstellungSchliessen := FALSE;
  steplWandverstellungOeffnen    := STEP_0_E;
  steplWandverstellungSchliessen := STEP_0_E;
  tonlEingefahrenWandEinlaufseite( IN := FALSE );
  tonlAusgefahrenWandEinlaufseite( IN := FALSE );
  tonlEingefahrenWandAuslaufseite( IN := FALSE );
  tonlAusgefahrenWandAuslaufseite( IN := FALSE );
  tonlBewegungszeitOeffnen( IN := FALSE );
  tonlBewegungszeitSchliessen( IN := FALSE );
  bpDone := FALSE;
ELSE
  WandverstellungOeffnen();
  WandverstellungSchliessen();
END_IF
END_FUNCTION_BLOCK
